  movel([0.339541, -0.797675, -2.797193, -1.117521, 1.570796, 1.910338],accel_mss,speed_ms,0,blend_radius_m)
  movel([0.338270, -0.798291, -2.797090, -1.117008, 1.570796, 1.909067],accel_mss,speed_ms,0,blend_radius_m)
  movel([0.337067, -0.798451, -2.797063, -1.116875, 1.570796, 1.907863],accel_mss,speed_ms,0,blend_radius_m)
  movel([0.336030, -0.798308, -2.797087, -1.116993, 1.570796, 1.906826],accel_mss,speed_ms,0,blend_radius_m)
  movel([0.330509, -0.796529, -2.797384, -1.118476, 1.570796, 1.901306],accel_mss,speed_ms,0,blend_radius_m)
  movel([0.325271, -0.794328, -2.797750, -1.120311, 1.570796, 1.896067],accel_mss,speed_ms,0,blend_radius_m)
  movel([0.320318, -0.791707, -2.798181, -1.122501, 1.570796, 1.891115],accel_mss,speed_ms,0,blend_radius_m)
  movel([0.315671, -0.788660, -2.798679, -1.125051, 1.570796, 1.886468],accel_mss,speed_ms,0,blend_radius_m)
  movel([0.314088, -0.787352, -2.798891, -1.126146, 1.570796, 1.884885],accel_mss,speed_ms,0,blend_radius_m)
  movel([0.312919, -0.785569, -2.799178, -1.127642, 1.570796, 1.883716],accel_mss,speed_ms,0,blend_radius_m)
  movel([0.312565, -0.784172, -2.799403, -1.128814, 1.570796, 1.883362],accel_mss,speed_ms,0,blend_radius_m)
  movel([0.312427, -0.782583, -2.799657, -1.130150, 1.570796, 1.883224],accel_mss,speed_ms,0,blend_radius_m)
  movel([0.312533, -0.779070, -2.800213, -1.133105, 1.570796, 1.883329],accel_mss,speed_ms,0,blend_radius_m)
  movel([0.314201, -0.765515, -2.802305, -1.144570, 1.570796, 1.884998],accel_mss,speed_ms,0,blend_radius_m)
  movel([0.314322, -0.761910, -2.802846, -1.147634, 1.570796, 1.885118],accel_mss,speed_ms,0,blend_radius_m)
  movel([0.313995, -0.758978, -2.803281, -1.150130, 1.570796, 1.884791],accel_mss,speed_ms,0,blend_radius_m)
  movel([0.313608, -0.757890, -2.803441, -1.151058, 1.570796, 1.884404],accel_mss,speed_ms,0,blend_radius_m)
  movel([0.313044, -0.757111, -2.803556, -1.151722, 1.570796, 1.883841],accel_mss,speed_ms,0,blend_radius_m)
  movel([0.312284, -0.756701, -2.803616, -1.152072, 1.570796, 1.883080],accel_mss,speed_ms,0,blend_radius_m)
  movel([0.311307, -0.756696, -2.803617, -1.152076, 1.570796, 1.882104],accel_mss,speed_ms,0,blend_radius_m)
  movel([0.309324, -0.757338, -2.803522, -1.151529, 1.570796, 1.880120],accel_mss,speed_ms,0,blend_radius_m)
  movel([0.308425, -0.757514, -2.803496, -1.151378, 1.570796, 1.879221],accel_mss,speed_ms,0,blend_radius_m)
  movel([0.307786, -0.757283, -2.803531, -1.151575, 1.570796, 1.878582],accel_mss,speed_ms,0,blend_radius_m)
  movel([0.307584, -0.756087, -2.803706, -1.152596, 1.570796, 1.878380],accel_mss,speed_ms,0,blend_radius_m)
  movel([0.307977, -0.754391, -2.803953, -1.154044, 1.570796, 1.878773],accel_mss,speed_ms,0,blend_radius_m)
  movel([0.309463, -0.748829, -2.804756, -1.158804, 1.570796, 1.880260],accel_mss,speed_ms,0,blend_radius_m)
  movel([0.310630, -0.743455, -2.805517, -1.163417, 1.570796, 1.881426],accel_mss,speed_ms,0,blend_radius_m)
  movel([0.312165, -0.733164, -2.806936, -1.172289, 1.570796, 1.882961],accel_mss,speed_ms,0,blend_radius_m)
  movel([0.312944, -0.723256, -2.808256, -1.180876, 1.570796, 1.883740],accel_mss,speed_ms,0,blend_radius_m)
  movel([0.313326, -0.713471, -2.809516, -1.189402, 1.570796, 1.884122],accel_mss,speed_ms,0,blend_radius_m)
  speed_ms = 0.005
  movel([0.313326, -0.706215, -2.802909, -1.203265, 1.570796, 1.884122],accel_mss,speed_ms,0,blend_radius_m)
  speed_ms = 0.040
  movel([0.305588, -0.724600, -2.800519, -1.187270, 1.570796, 1.876385],accel_mss,speed_ms,0,blend_radius_m)
  speed_ms = 0.005
  movel([0.305588, -0.732101, -2.807080, -1.173208, 1.570796, 1.876385],accel_mss,speed_ms,0,blend_radius_m)
  speed_ms = 0.025
  movel([0.301170, -0.744287, -2.805400, -1.162703, 1.570796, 1.871966],accel_mss,speed_ms,0,blend_radius_m)
  movel([0.298692, -0.750428, -2.804526, -1.157434, 1.570796, 1.869489],accel_mss,speed_ms,0,blend_radius_m)
  movel([0.296052, -0.756579, -2.803634, -1.152176, 1.570796, 1.866849],accel_mss,speed_ms,0,blend_radius_m)
  movel([0.293909, -0.755261, -2.803827, -1.153301, 1.570796, 1.864706],accel_mss,speed_ms,0,blend_radius_m)
  movel([0.293492, -0.755110, -2.803849, -1.153430, 1.570796, 1.864289],accel_mss,speed_ms,0,blend_radius_m)
  movel([0.292925, -0.755314, -2.803819, -1.153256, 1.570796, 1.863721],accel_mss,speed_ms,0,blend_radius_m)
  movel([0.292315, -0.755987, -2.803720, -1.152681, 1.570796, 1.863111],accel_mss,speed_ms,0,blend_radius_m)
  movel([0.291839, -0.756807, -2.803600, -1.151981, 1.570796, 1.862635],accel_mss,speed_ms,0,blend_radius_m)
  movel([0.288894, -0.761863, -2.802853, -1.147674, 1.570796, 1.859691],accel_mss,speed_ms,0,blend_radius_m)
  movel([0.285493, -0.766786, -2.802112, -1.143491, 1.570796, 1.856290],accel_mss,speed_ms,0,blend_radius_m)
  movel([0.284595, -0.767854, -2.801950, -1.142584, 1.570796, 1.855391],accel_mss,speed_ms,0,blend_radius_m)
  movel([0.283710, -0.768447, -2.801860, -1.142082, 1.570796, 1.854506],accel_mss,speed_ms,0,blend_radius_m)
  movel([0.283279, -0.768196, -2.801898, -1.142295, 1.570796, 1.854075],accel_mss,speed_ms,0,blend_radius_m)
  movel([0.283199, -0.767514, -2.802002, -1.142873, 1.570796, 1.853995],accel_mss,speed_ms,0,blend_radius_m)
  movel([0.283611, -0.762679, -2.802731, -1.146980, 1.570796, 1.854408],accel_mss,speed_ms,0,blend_radius_m)
  movel([0.284807, -0.757324, -2.803525, -1.151541, 1.570796, 1.855604],accel_mss,speed_ms,0,blend_radius_m)
  speed_ms = 0.005
  movel([0.284807, -0.749511, -2.797028, -1.165850, 1.570796, 1.855604],accel_mss,speed_ms,0,blend_radius_m)
  speed_ms = 0.040
  movel([0.290706, -0.756584, -2.795983, -1.159821, 1.570796, 1.861503],accel_mss,speed_ms,0,blend_radius_m)
  speed_ms = 0.005
  movel([0.290706, -0.764482, -2.802460, -1.145446, 1.570796, 1.861503],accel_mss,speed_ms,0,blend_radius_m)
  speed_ms = 0.025
  movel([0.289009, -0.772297, -2.801270, -1.138822, 1.570796, 1.859805],accel_mss,speed_ms,0,blend_radius_m)
  movel([0.287811, -0.776370, -2.800637, -1.135382, 1.570796, 1.858608],accel_mss,speed_ms,0,blend_radius_m)
  movel([0.284778, -0.784728, -2.799313, -1.128347, 1.570796, 1.855575],accel_mss,speed_ms,0,blend_radius_m)
  movel([0.282956, -0.788978, -2.798627, -1.124784, 1.570796, 1.853753],accel_mss,speed_ms,0,blend_radius_m)
  movel([0.278747, -0.797523, -2.797219, -1.117648, 1.570796, 1.849544],accel_mss,speed_ms,0,blend_radius_m)
  movel([0.279478, -0.794879, -2.797658, -1.119852, 1.570796, 1.850275],accel_mss,speed_ms,0,blend_radius_m)
  movel([0.279565, -0.792616, -2.798032, -1.121741, 1.570796, 1.850361],accel_mss,speed_ms,0,blend_radius_m)
  movel([0.279016, -0.790889, -2.798315, -1.123185, 1.570796, 1.849813],accel_mss,speed_ms,0,blend_radius_m)
  movel([0.277841, -0.789851, -2.798485, -1.124053, 1.570796, 1.848637],accel_mss,speed_ms,0,blend_radius_m)
  speed_ms = 0.005
  movel([0.277841, -0.781667, -2.792079, -1.138643, 1.570796, 1.848637],accel_mss,speed_ms,0,blend_radius_m)
  speed_ms = 0.040
  movel([0.251919, -0.798788, -2.789231, -1.124370, 1.570796, 1.822716],accel_mss,speed_ms,0,blend_radius_m)
  speed_ms = 0.005
  movel([0.251919, -0.807155, -2.795586, -1.109648, 1.570796, 1.822716],accel_mss,speed_ms,0,blend_radius_m)
  speed_ms = 0.025
  movel([0.247378, -0.813004, -2.794571, -1.104814, 1.570796, 1.818174],accel_mss,speed_ms,0,blend_radius_m)
  movel([0.242549, -0.818489, -2.793603, -1.100297, 1.570796, 1.813345],accel_mss,speed_ms,0,blend_radius_m)
  movel([0.237519, -0.823531, -2.792698, -1.096159, 1.570796, 1.808315],accel_mss,speed_ms,0,blend_radius_m)
  movel([0.232368, -0.828046, -2.791877, -1.092466, 1.570796, 1.803164],accel_mss,speed_ms,0,blend_radius_m)
  movel([0.233688, -0.825444, -2.792352, -1.094593, 1.570796, 1.804484],accel_mss,speed_ms,0,blend_radius_m)
  movel([0.234683, -0.823023, -2.792790, -1.096576, 1.570796, 1.805479],accel_mss,speed_ms,0,blend_radius_m)
  movel([0.235280, -0.821000, -2.793154, -1.098235, 1.570796, 1.806076],accel_mss,speed_ms,0,blend_radius_m)
  movel([0.235407, -0.819588, -2.793407, -1.099394, 1.570796, 1.806203],accel_mss,speed_ms,0,blend_radius_m)
  movel([0.234984, -0.819018, -2.793509, -1.099863, 1.570796, 1.805780],accel_mss,speed_ms,0,blend_radius_m)
  movel([0.234547, -0.819112, -2.793492, -1.099785, 1.570796, 1.805344],accel_mss,speed_ms,0,blend_radius_m)
  movel([0.233940, -0.819499, -2.793423, -1.099468, 1.570796, 1.804736],accel_mss,speed_ms,0,blend_radius_m)
  movel([0.232209, -0.821250, -2.793109, -1.098030, 1.570796, 1.803005],accel_mss,speed_ms,0,blend_radius_m)
  movel([0.227802, -0.827037, -2.792062, -1.093291, 1.570796, 1.798598],accel_mss,speed_ms,0,blend_radius_m)
  movel([0.225752, -0.829544, -2.791602, -1.091243, 1.570796, 1.796549],accel_mss,speed_ms,0,blend_radius_m)
  movel([0.221376, -0.834255, -2.790729, -1.087405, 1.570796, 1.792172],accel_mss,speed_ms,0,blend_radius_m)
  movel([0.219102, -0.836398, -2.790328, -1.085663, 1.570796, 1.789898],accel_mss,speed_ms,0,blend_radius_m)
  movel([0.216804, -0.838351, -2.789960, -1.084077, 1.570796, 1.787600],accel_mss,speed_ms,0,blend_radius_m)
  movel([0.214506, -0.840095, -2.789630, -1.082663, 1.570796, 1.785302],accel_mss,speed_ms,0,blend_radius_m)
  movel([0.212240, -0.841584, -2.789347, -1.081458, 1.570796, 1.783037],accel_mss,speed_ms,0,blend_radius_m)
  movel([0.215104, -0.837462, -2.790128, -1.084799, 1.570796, 1.785901],accel_mss,speed_ms,0,blend_radius_m)
  movel([0.217906, -0.833284, -2.790910, -1.088195, 1.570796, 1.788702],accel_mss,speed_ms,0,blend_radius_m)
  movel([0.219209, -0.830564, -2.791414, -1.090411, 1.570796, 1.790005],accel_mss,speed_ms,0,blend_radius_m)
  movel([0.219966, -0.827999, -2.791886, -1.092505, 1.570796, 1.790763],accel_mss,speed_ms,0,blend_radius_m)
  movel([0.219920, -0.827191, -2.792033, -1.093165, 1.570796, 1.790716],accel_mss,speed_ms,0,blend_radius_m)
  movel([0.219466, -0.826927, -2.792082, -1.093380, 1.570796, 1.790262],accel_mss,speed_ms,0,blend_radius_m)
  movel([0.218525, -0.827372, -2.792000, -1.093017, 1.570796, 1.789321],accel_mss,speed_ms,0,blend_radius_m)
  movel([0.217006, -0.828695, -2.791758, -1.091936, 1.570796, 1.787803],accel_mss,speed_ms,0,blend_radius_m)
  movel([0.209003, -0.836814, -2.790250, -1.085325, 1.570796, 1.779799],accel_mss,speed_ms,0,blend_radius_m)
  movel([0.205006, -0.840380, -2.789576, -1.082433, 1.570796, 1.775803],accel_mss,speed_ms,0,blend_radius_m)
  movel([0.203015, -0.841850, -2.789296, -1.081243, 1.570796, 1.773811],accel_mss,speed_ms,0,blend_radius_m)
  movel([0.201023, -0.843044, -2.789068, -1.080276, 1.570796, 1.771819],accel_mss,speed_ms,0,blend_radius_m)
  speed_ms = 0.005
  movel([0.201023, -0.834334, -2.782823, -1.095231, 1.570796, 1.771819],accel_mss,speed_ms,0,blend_radius_m)
  speed_ms = 0.040
  movel([0.238662, -0.779480, -2.792432, -1.140477, 1.570796, 1.809458],accel_mss,speed_ms,0,blend_radius_m)
  speed_ms = 0.005
  movel([0.238662, -0.787640, -2.798844, -1.125905, 1.570796, 1.809458],accel_mss,speed_ms,0,blend_radius_m)
  speed_ms = 0.025
  movel([0.238890, -0.784551, -2.799342, -1.128496, 1.570796, 1.809686],accel_mss,speed_ms,0,blend_radius_m)
  movel([0.239732, -0.781111, -2.799891, -1.131387, 1.570796, 1.810528],accel_mss,speed_ms,0,blend_radius_m)
  movel([0.241121, -0.777396, -2.800477, -1.134517, 1.570796, 1.811917],accel_mss,speed_ms,0,blend_radius_m)
  movel([0.242984, -0.773502, -2.801083, -1.137804, 1.570796, 1.813781],accel_mss,speed_ms,0,blend_radius_m)
  movel([0.245268, -0.769501, -2.801699, -1.141189, 1.570796, 1.816064],accel_mss,speed_ms,0,blend_radius_m)
  movel([0.247890, -0.765497, -2.802307, -1.144584, 1.570796, 1.818687],accel_mss,speed_ms,0,blend_radius_m)
  movel([0.250794, -0.761568, -2.802896, -1.147924, 1.570796, 1.821590],accel_mss,speed_ms,0,blend_radius_m)
  movel([0.253896, -0.757818, -2.803452, -1.151119, 1.570796, 1.824692],accel_mss,speed_ms,0,blend_radius_m)
  movel([0.257898, -0.753459, -2.804089, -1.154841, 1.570796, 1.828695],accel_mss,speed_ms,0,blend_radius_m)
  movel([0.266086, -0.744895, -2.805314, -1.162180, 1.570796, 1.836882],accel_mss,speed_ms,0,blend_radius_m)
  movel([0.270058, -0.740350, -2.805950, -1.166089, 1.570796, 1.840855],accel_mss,speed_ms,0,blend_radius_m)
  movel([0.273771, -0.735350, -2.806639, -1.170400, 1.570796, 1.844568],accel_mss,speed_ms,0,blend_radius_m)
  movel([0.275420, -0.732740, -2.806993, -1.172655, 1.570796, 1.846216],accel_mss,speed_ms,0,blend_radius_m)
  movel([0.276854, -0.730144, -2.807343, -1.174902, 1.570796, 1.847650],accel_mss,speed_ms,0,blend_radius_m)
  movel([0.278016, -0.727626, -2.807680, -1.177084, 1.570796, 1.848812],accel_mss,speed_ms,0,blend_radius_m)
  movel([0.278854, -0.725248, -2.807995, -1.179146, 1.570796, 1.849650],accel_mss,speed_ms,0,blend_radius_m)
  movel([0.279296, -0.723094, -2.808277, -1.181017, 1.570796, 1.850092],accel_mss,speed_ms,0,blend_radius_m)
  movel([0.279283, -0.721232, -2.808520, -1.182636, 1.570796, 1.850080],accel_mss,speed_ms,0,blend_radius_m)
  speed_ms = 0.005
  movel([0.279283, -0.713873, -2.801932, -1.196584, 1.570796, 1.850080],accel_mss,speed_ms,0,blend_radius_m)
  speed_ms = 0.040
  movel([0.278218, -0.699673, -2.803723, -1.208993, 1.570796, 1.849015],accel_mss,speed_ms,0,blend_radius_m)
  speed_ms = 0.005
  movel([0.278218, -0.706840, -2.810345, -1.195204, 1.570796, 1.849015],accel_mss,speed_ms,0,blend_radius_m)
  speed_ms = 0.025
  movel([0.274128, -0.720252, -2.808648, -1.183489, 1.570796, 1.844925],accel_mss,speed_ms,0,blend_radius_m)
  movel([0.272708, -0.723399, -2.808238, -1.180753, 1.570796, 1.843504],accel_mss,speed_ms,0,blend_radius_m)
  movel([0.270637, -0.726538, -2.807824, -1.178027, 1.570796, 1.841433],accel_mss,speed_ms,0,blend_radius_m)
  movel([0.268156, -0.729467, -2.807434, -1.175488, 1.570796, 1.838952],accel_mss,speed_ms,0,blend_radius_m)
  movel([0.259858, -0.738116, -2.806259, -1.168014, 1.570796, 1.830654],accel_mss,speed_ms,0,blend_radius_m)
  movel([0.257055, -0.741410, -2.805803, -1.165176, 1.570796, 1.827852],accel_mss,speed_ms,0,blend_radius_m)
  movel([0.254399, -0.744824, -2.805324, -1.162241, 1.570796, 1.825196],accel_mss,speed_ms,0,blend_radius_m)
  movel([0.251913, -0.748315, -2.804829, -1.159245, 1.570796, 1.822709],accel_mss,speed_ms,0,blend_radius_m)
  movel([0.249806, -0.751776, -2.804332, -1.156281, 1.570796, 1.820602],accel_mss,speed_ms,0,blend_radius_m)
  movel([0.248006, -0.755228, -2.803831, -1.153329, 1.570796, 1.818802],accel_mss,speed_ms,0,blend_radius_m)
  movel([0.246241, -0.758651, -2.803329, -1.150409, 1.570796, 1.817038],accel_mss,speed_ms,0,blend_radius_m)
  movel([0.244246, -0.762033, -2.802827, -1.147529, 1.570796, 1.815042],accel_mss,speed_ms,0,blend_radius_m)
  movel([0.242758, -0.756334, -2.803670, -1.152385, 1.570796, 1.813555],accel_mss,speed_ms,0,blend_radius_m)
  movel([0.243050, -0.754319, -2.803964, -1.154106, 1.570796, 1.813846],accel_mss,speed_ms,0,blend_radius_m)
  movel([0.243651, -0.752175, -2.804275, -1.155940, 1.570796, 1.814448],accel_mss,speed_ms,0,blend_radius_m)
  movel([0.244562, -0.749898, -2.804603, -1.157888, 1.570796, 1.815359],accel_mss,speed_ms,0,blend_radius_m)
  movel([0.245801, -0.747468, -2.804950, -1.159971, 1.570796, 1.816598],accel_mss,speed_ms,0,blend_radius_m)
  movel([0.248098, -0.744058, -2.805432, -1.162899, 1.570796, 1.818894],accel_mss,speed_ms,0,blend_radius_m)
  movel([0.251441, -0.739885, -2.806015, -1.166489, 1.570796, 1.822238],accel_mss,speed_ms,0,blend_radius_m)
  movel([0.259675, -0.730420, -2.807306, -1.174663, 1.570796, 1.830471],accel_mss,speed_ms,0,blend_radius_m)
  movel([0.263755, -0.725728, -2.807931, -1.178730, 1.570796, 1.834551],accel_mss,speed_ms,0,blend_radius_m)
  movel([0.267253, -0.721467, -2.808490, -1.182432, 1.570796, 1.838049],accel_mss,speed_ms,0,blend_radius_m)
  movel([0.269743, -0.717961, -2.808943, -1.185485, 1.570796, 1.840539],accel_mss,speed_ms,0,blend_radius_m)
  movel([0.270479, -0.716582, -2.809120, -1.186687, 1.570796, 1.841275],accel_mss,speed_ms,0,blend_radius_m)
  movel([0.270799, -0.715510, -2.809257, -1.187622, 1.570796, 1.841595],accel_mss,speed_ms,0,blend_radius_m)
  speed_ms = 0.005
  movel([0.270799, -0.708226, -2.802655, -1.201508, 1.570796, 1.841595],accel_mss,speed_ms,0,blend_radius_m)
  speed_ms = 0.040
  movel([0.256086, -0.711101, -2.802289, -1.198999, 1.570796, 1.826882],accel_mss,speed_ms,0,blend_radius_m)
  speed_ms = 0.005
  movel([0.256086, -0.718423, -2.808884, -1.185082, 1.570796, 1.826882],accel_mss,speed_ms,0,blend_radius_m)
  speed_ms = 0.025
  movel([0.254666, -0.718676, -2.808851, -1.184862, 1.570796, 1.825462],accel_mss,speed_ms,0,blend_radius_m)
  movel([0.253508, -0.718501, -2.808874, -1.185014, 1.570796, 1.824304],accel_mss,speed_ms,0,blend_radius_m)
  movel([0.251855, -0.717143, -2.809048, -1.186198, 1.570796, 1.822651],accel_mss,speed_ms,0,blend_radius_m)
  movel([0.250882, -0.714842, -2.809342, -1.188205, 1.570796, 1.821679],accel_mss,speed_ms,0,blend_radius_m)
  movel([0.250362, -0.712082, -2.809691, -1.190616, 1.570796, 1.821158],accel_mss,speed_ms,0,blend_radius_m)
  movel([0.250376, -0.710916, -2.809838, -1.191635, 1.570796, 1.821172],accel_mss,speed_ms,0,blend_radius_m)
  movel([0.251431, -0.708572, -2.810131, -1.193686, 1.570796, 1.822227],accel_mss,speed_ms,0,blend_radius_m)
  movel([0.255097, -0.701778, -2.810965, -1.199646, 1.570796, 1.825893],accel_mss,speed_ms,0,blend_radius_m)
  movel([0.261993, -0.688097, -2.812584, -1.211708, 1.570796, 1.832789],accel_mss,speed_ms,0,blend_radius_m)
  movel([0.265206, -0.681243, -2.813364, -1.217782, 1.570796, 1.836002],accel_mss,speed_ms,0,blend_radius_m)
  speed_ms = 0.005
  movel([0.265206, -0.674435, -2.806684, -1.231270, 1.570796, 1.836002],accel_mss,speed_ms,0,blend_radius_m)
  speed_ms = 0.040
  movel([0.255172, -0.681907, -2.805837, -1.224645, 1.570796, 1.825968],accel_mss,speed_ms,0,blend_radius_m)
  speed_ms = 0.005
  movel([0.255172, -0.688824, -2.812500, -1.211066, 1.570796, 1.825968],accel_mss,speed_ms,0,blend_radius_m)
  speed_ms = 0.025
  movel([0.253576, -0.692842, -2.812032, -1.207515, 1.570796, 1.824373],accel_mss,speed_ms,0,blend_radius_m)
  movel([0.251612, -0.696958, -2.811545, -1.203886, 1.570796, 1.822409],accel_mss,speed_ms,0,blend_radius_m)
  movel([0.249200, -0.700991, -2.811060, -1.200338, 1.570796, 1.819996],accel_mss,speed_ms,0,blend_radius_m)
  movel([0.247798, -0.702929, -2.810825, -1.198635, 1.570796, 1.818594],accel_mss,speed_ms,0,blend_radius_m)
  movel([0.244762, -0.706607, -2.810374, -1.195408, 1.570796, 1.815558],accel_mss,speed_ms,0,blend_radius_m)
  movel([0.243999, -0.708241, -2.810172, -1.193976, 1.570796, 1.814795],accel_mss,speed_ms,0,blend_radius_m)
  movel([0.239388, -0.720425, -2.808625, -1.183339, 1.570796, 1.810184],accel_mss,speed_ms,0,blend_radius_m)
  movel([0.238976, -0.721588, -2.808474, -1.182327, 1.570796, 1.809772],accel_mss,speed_ms,0,blend_radius_m)
  movel([0.238840, -0.722571, -2.808346, -1.181472, 1.570796, 1.809637],accel_mss,speed_ms,0,blend_radius_m)
  movel([0.239436, -0.723273, -2.808254, -1.180862, 1.570796, 1.810232],accel_mss,speed_ms,0,blend_radius_m)
  movel([0.240542, -0.723333, -2.808246, -1.180810, 1.570796, 1.811338],accel_mss,speed_ms,0,blend_radius_m)
  movel([0.243805, -0.723330, -2.808247, -1.180812, 1.570796, 1.814601],accel_mss,speed_ms,0,blend_radius_m)
  movel([0.246751, -0.723842, -2.808179, -1.180368, 1.570796, 1.817547],accel_mss,speed_ms,0,blend_radius_m)
  movel([0.249147, -0.725096, -2.808014, -1.179278, 1.570796, 1.819943],accel_mss,speed_ms,0,blend_radius_m)
  movel([0.250740, -0.727339, -2.807718, -1.177332, 1.570796, 1.821537],accel_mss,speed_ms,0,blend_radius_m)
  speed_ms = 0.005
  movel([0.250740, -0.719899, -2.801145, -1.191345, 1.570796, 1.821537],accel_mss,speed_ms,0,blend_radius_m)
  speed_ms = 0.040
  movel([0.239180, -0.750332, -2.796908, -1.165149, 1.570796, 1.809976],accel_mss,speed_ms,0,blend_radius_m)
  speed_ms = 0.005
  movel([0.239180, -0.758155, -2.803402, -1.150831, 1.570796, 1.809976],accel_mss,speed_ms,0,blend_radius_m)
  speed_ms = 0.025
  movel([0.238467, -0.758887, -2.803294, -1.150207, 1.570796, 1.809264],accel_mss,speed_ms,0,blend_radius_m)
  movel([0.237810, -0.759796, -2.803160, -1.149434, 1.570796, 1.808607],accel_mss,speed_ms,0,blend_radius_m)
  movel([0.235162, -0.764438, -2.802467, -1.145484, 1.570796, 1.805958],accel_mss,speed_ms,0,blend_radius_m)
  movel([0.234732, -0.764883, -2.802400, -1.145106, 1.570796, 1.805529],accel_mss,speed_ms,0,blend_radius_m)
  movel([0.234120, -0.765111, -2.802365, -1.144913, 1.570796, 1.804916],accel_mss,speed_ms,0,blend_radius_m)
  movel([0.233671, -0.764874, -2.802401, -1.145114, 1.570796, 1.804467],accel_mss,speed_ms,0,blend_radius_m)
  movel([0.233188, -0.763476, -2.802611, -1.146302, 1.570796, 1.803984],accel_mss,speed_ms,0,blend_radius_m)
  movel([0.233194, -0.760208, -2.803099, -1.149082, 1.570796, 1.803991],accel_mss,speed_ms,0,blend_radius_m)
  movel([0.234136, -0.756594, -2.803632, -1.152163, 1.570796, 1.804933],accel_mss,speed_ms,0,blend_radius_m)
  movel([0.235569, -0.752720, -2.804196, -1.155473, 1.570796, 1.806365],accel_mss,speed_ms,0,blend_radius_m)
  movel([0.237248, -0.748804, -2.804759, -1.158826, 1.570796, 1.808045],accel_mss,speed_ms,0,blend_radius_m)
  movel([0.239202, -0.744941, -2.805308, -1.162141, 1.570796, 1.809999],accel_mss,speed_ms,0,blend_radius_m)
  movel([0.241419, -0.741136, -2.805841, -1.165412, 1.570796, 1.812215],accel_mss,speed_ms,0,blend_radius_m)
  movel([0.243887, -0.737388, -2.806360, -1.168642, 1.570796, 1.814683],accel_mss,speed_ms,0,blend_radius_m)
  movel([0.246599, -0.733692, -2.806864, -1.171832, 1.570796, 1.817396],accel_mss,speed_ms,0,blend_radius_m)
  movel([0.249538, -0.730058, -2.807355, -1.174976, 1.570796, 1.820334],accel_mss,speed_ms,0,blend_radius_m)
  movel([0.252702, -0.726473, -2.807833, -1.178083, 1.570796, 1.823499],accel_mss,speed_ms,0,blend_radius_m)
  movel([0.256073, -0.722947, -2.808297, -1.181146, 1.570796, 1.826870],accel_mss,speed_ms,0,blend_radius_m)
  movel([0.260755, -0.717676, -2.808980, -1.185733, 1.570796, 1.831551],accel_mss,speed_ms,0,blend_radius_m)
  movel([0.265685, -0.711492, -2.809766, -1.191132, 1.570796, 1.836482],accel_mss,speed_ms,0,blend_radius_m)
  movel([0.271037, -0.704320, -2.810655, -1.197413, 1.570796, 1.841833],accel_mss,speed_ms,0,blend_radius_m)
  speed_ms = 0.005
  movel([0.271037, -0.697188, -2.804027, -1.211174, 1.570796, 1.841833],accel_mss,speed_ms,0,blend_radius_m)
  speed_ms = 0.040
  movel([0.266633, -0.698799, -2.803830, -1.209760, 1.570796, 1.837429],accel_mss,speed_ms,0,blend_radius_m)
  speed_ms = 0.005
  movel([0.266633, -0.705953, -2.810455, -1.195981, 1.570796, 1.837429],accel_mss,speed_ms,0,blend_radius_m)
  speed_ms = 0.025
  movel([0.271058, -0.696231, -2.811631, -1.204527, 1.570796, 1.841854],accel_mss,speed_ms,0,blend_radius_m)
  movel([0.275991, -0.686298, -2.812790, -1.213301, 1.570796, 1.846787],accel_mss,speed_ms,0,blend_radius_m)
  movel([0.278750, -0.681294, -2.813358, -1.217737, 1.570796, 1.849546],accel_mss,speed_ms,0,blend_radius_m)
  movel([0.281743, -0.676290, -2.813915, -1.222183, 1.570796, 1.852540],accel_mss,speed_ms,0,blend_radius_m)
  movel([0.285025, -0.671298, -2.814460, -1.226631, 1.570796, 1.855822],accel_mss,speed_ms,0,blend_radius_m)
  movel([0.288616, -0.666352, -2.814990, -1.231047, 1.570796, 1.859412],accel_mss,speed_ms,0,blend_radius_m)
  movel([0.298570, -0.653944, -2.816274, -1.242171, 1.570796, 1.869366],accel_mss,speed_ms,0,blend_radius_m)
  movel([0.302903, -0.648242, -2.816842, -1.247305, 1.570796, 1.873699],accel_mss,speed_ms,0,blend_radius_m)
  movel([0.304959, -0.645315, -2.817129, -1.249945, 1.570796, 1.875755],accel_mss,speed_ms,0,blend_radius_m)
  movel([0.306841, -0.642327, -2.817418, -1.252645, 1.570796, 1.877638],accel_mss,speed_ms,0,blend_radius_m)
  movel([0.311183, -0.633365, -2.818263, -1.260761, 1.570796, 1.881979],accel_mss,speed_ms,0,blend_radius_m)
  speed_ms = 0.005
  movel([0.311183, -0.627283, -2.811487, -1.273619, 1.570796, 1.881979],accel_mss,speed_ms,0,blend_radius_m)
  speed_ms = 0.040
  movel([0.321759, -0.606621, -2.813304, -1.292463, 1.570796, 1.892555],accel_mss,speed_ms,0,blend_radius_m)
  speed_ms = 0.005
  movel([0.321759, -0.612365, -2.820117, -1.279907, 1.570796, 1.892555],accel_mss,speed_ms,0,blend_radius_m)
  speed_ms = 0.025
  movel([0.325188, -0.604942, -2.820730, -1.286716, 1.570796, 1.895984],accel_mss,speed_ms,0,blend_radius_m)
  movel([0.327388, -0.601192, -2.821032, -1.290165, 1.570796, 1.898185],accel_mss,speed_ms,0,blend_radius_m)
  movel([0.330084, -0.597532, -2.821322, -1.293535, 1.570796, 1.900880],accel_mss,speed_ms,0,blend_radius_m)
  movel([0.332238, -0.595164, -2.821506, -1.295719, 1.570796, 1.903034],accel_mss,speed_ms,0,blend_radius_m)
  movel([0.334479, -0.593024, -2.821671, -1.297694, 1.570796, 1.905275],accel_mss,speed_ms,0,blend_radius_m)
  movel([0.339064, -0.589097, -2.821969, -1.301323, 1.570796, 1.909861],accel_mss,speed_ms,0,blend_radius_m)
  movel([0.343198, -0.585241, -2.822256, -1.304892, 1.570796, 1.913994],accel_mss,speed_ms,0,blend_radius_m)
  movel([0.346574, -0.581375, -2.822538, -1.308476, 1.570796, 1.917370],accel_mss,speed_ms,0,blend_radius_m)
  movel([0.353165, -0.572343, -2.823174, -1.316871, 1.570796, 1.923961],accel_mss,speed_ms,0,blend_radius_m)
  movel([0.354587, -0.570547, -2.823297, -1.318544, 1.570796, 1.925383],accel_mss,speed_ms,0,blend_radius_m)
  movel([0.356113, -0.568928, -2.823407, -1.320054, 1.570796, 1.926909],accel_mss,speed_ms,0,blend_radius_m)
  movel([0.359378, -0.566081, -2.823598, -1.322710, 1.570796, 1.930174],accel_mss,speed_ms,0,blend_radius_m)
  movel([0.365995, -0.560955, -2.823934, -1.327500, 1.570796, 1.936792],accel_mss,speed_ms,0,blend_radius_m)
  movel([0.373073, -0.554833, -2.824322, -1.333234, 1.570796, 1.943869],accel_mss,speed_ms,0,blend_radius_m)
  movel([0.376615, -0.551458, -2.824530, -1.336401, 1.570796, 1.947411],accel_mss,speed_ms,0,blend_radius_m)
  movel([0.380090, -0.547720, -2.824756, -1.339913, 1.570796, 1.950886],accel_mss,speed_ms,0,blend_radius_m)
  movel([0.382697, -0.544354, -2.824954, -1.343081, 1.570796, 1.953493],accel_mss,speed_ms,0,blend_radius_m)
  movel([0.384821, -0.540887, -2.825155, -1.346348, 1.570796, 1.955617],accel_mss,speed_ms,0,blend_radius_m)
  movel([0.385968, -0.537961, -2.825321, -1.349107, 1.570796, 1.956764],accel_mss,speed_ms,0,blend_radius_m)
  movel([0.386018, -0.536910, -2.825379, -1.350100, 1.570796, 1.956814],accel_mss,speed_ms,0,blend_radius_m)
  movel([0.385633, -0.536242, -2.825417, -1.350731, 1.570796, 1.956430],accel_mss,speed_ms,0,blend_radius_m)
  movel([0.384024, -0.535820, -2.825440, -1.351129, 1.570796, 1.954820],accel_mss,speed_ms,0,blend_radius_m)
  movel([0.381703, -0.536196, -2.825419, -1.350773, 1.570796, 1.952500],accel_mss,speed_ms,0,blend_radius_m)
  movel([0.378837, -0.537272, -2.825359, -1.349758, 1.570796, 1.949633],accel_mss,speed_ms,0,blend_radius_m)
  movel([0.375629, -0.538907, -2.825267, -1.348215, 1.570796, 1.946425],accel_mss,speed_ms,0,blend_radius_m)
  movel([0.372254, -0.541002, -2.825148, -1.346239, 1.570796, 1.943051],accel_mss,speed_ms,0,blend_radius_m)
  movel([0.368906, -0.543422, -2.825009, -1.343959, 1.570796, 1.939702],accel_mss,speed_ms,0,blend_radius_m)
  movel([0.365765, -0.546056, -2.824854, -1.341478, 1.570796, 1.936562],accel_mss,speed_ms,0,blend_radius_m)
  movel([0.363011, -0.548786, -2.824692, -1.338911, 1.570796, 1.933807],accel_mss,speed_ms,0,blend_radius_m)
  movel([0.359228, -0.553381, -2.824412, -1.334596, 1.570796, 1.930024],accel_mss,speed_ms,0,blend_radius_m)
  movel([0.348676, -0.567496, -2.823503, -1.321389, 1.570796, 1.919472],accel_mss,speed_ms,0,blend_radius_m)
  movel([0.341420, -0.576528, -2.822883, -1.312977, 1.570796, 1.912216],accel_mss,speed_ms,0,blend_radius_m)
  movel([0.334837, -0.583796, -2.822362, -1.306231, 1.570796, 1.905633],accel_mss,speed_ms,0,blend_radius_m)
  movel([0.331585, -0.587318, -2.822102, -1.302969, 1.570796, 1.902381],accel_mss,speed_ms,0,blend_radius_m)
  movel([0.328499, -0.590976, -2.821827, -1.299586, 1.570796, 1.899296],accel_mss,speed_ms,0,blend_radius_m)
  movel([0.325566, -0.594946, -2.821523, -1.295920, 1.570796, 1.896362],accel_mss,speed_ms,0,blend_radius_m)
  movel([0.322921, -0.598937, -2.821211, -1.292241, 1.570796, 1.893717],accel_mss,speed_ms,0,blend_radius_m)
  movel([0.320533, -0.602936, -2.820893, -1.288561, 1.570796, 1.891330],accel_mss,speed_ms,0,blend_radius_m)
  movel([0.318373, -0.606911, -2.820570, -1.284908, 1.570796, 1.889170],accel_mss,speed_ms,0,blend_radius_m)
  movel([0.314600, -0.614729, -2.819917, -1.277743, 1.570796, 1.885397],accel_mss,speed_ms,0,blend_radius_m)
  movel([0.311326, -0.622247, -2.819266, -1.270876, 1.570796, 1.882122],accel_mss,speed_ms,0,blend_radius_m)
  speed_ms = 0.005
  movel([0.311326, -0.616343, -2.812471, -1.283575, 1.570796, 1.882122],accel_mss,speed_ms,0,blend_radius_m)
  speed_ms = 0.040
  movel([0.303174, -0.623517, -2.811831, -1.277041, 1.570796, 1.873970],accel_mss,speed_ms,0,blend_radius_m)
  speed_ms = 0.005
  movel([0.303174, -0.629538, -2.818614, -1.264237, 1.570796, 1.873970],accel_mss,speed_ms,0,blend_radius_m)
  speed_ms = 0.025
  movel([0.308567, -0.617650, -2.819667, -1.275073, 1.570796, 1.879363],accel_mss,speed_ms,0,blend_radius_m)
  movel([0.311017, -0.612601, -2.820097, -1.279692, 1.570796, 1.881813],accel_mss,speed_ms,0,blend_radius_m)
  movel([0.313262, -0.607608, -2.820512, -1.284269, 1.570796, 1.884058],accel_mss,speed_ms,0,blend_radius_m)
  movel([0.314771, -0.603470, -2.820849, -1.288069, 1.570796, 1.885567],accel_mss,speed_ms,0,blend_radius_m)
  movel([0.315798, -0.599597, -2.821159, -1.291633, 1.570796, 1.886594],accel_mss,speed_ms,0,blend_radius_m)
  movel([0.316319, -0.596066, -2.821436, -1.294887, 1.570796, 1.887116],accel_mss,speed_ms,0,blend_radius_m)
  movel([0.316316, -0.592963, -2.821676, -1.297751, 1.570796, 1.887112],accel_mss,speed_ms,0,blend_radius_m)
  movel([0.318007, -0.591634, -2.821777, -1.298978, 1.570796, 1.888803],accel_mss,speed_ms,0,blend_radius_m)
  movel([0.319623, -0.590705, -2.821848, -1.299836, 1.570796, 1.890419],accel_mss,speed_ms,0,blend_radius_m)
  movel([0.322733, -0.589352, -2.821950, -1.301087, 1.570796, 1.893529],accel_mss,speed_ms,0,blend_radius_m)
  movel([0.326035, -0.587632, -2.822079, -1.302678, 1.570796, 1.896831],accel_mss,speed_ms,0,blend_radius_m)
  movel([0.327738, -0.586341, -2.822175, -1.303874, 1.570796, 1.898535],accel_mss,speed_ms,0,blend_radius_m)
  movel([0.329386, -0.584617, -2.822302, -1.305470, 1.570796, 1.900182],accel_mss,speed_ms,0,blend_radius_m)
  movel([0.348272, -0.561777, -2.823880, -1.326732, 1.570796, 1.919069],accel_mss,speed_ms,0,blend_radius_m)
  movel([0.348583, -0.559341, -2.824037, -1.329011, 1.570796, 1.919380],accel_mss,speed_ms,0,blend_radius_m)
  movel([0.348124, -0.557514, -2.824154, -1.330722, 1.570796, 1.918921],accel_mss,speed_ms,0,blend_radius_m)
  movel([0.346919, -0.556394, -2.824224, -1.331771, 1.570796, 1.917716],accel_mss,speed_ms,0,blend_radius_m)
  movel([0.345019, -0.556063, -2.824245, -1.332082, 1.570796, 1.915815],accel_mss,speed_ms,0,blend_radius_m)
  movel([0.348929, -0.553661, -2.824395, -1.334333, 1.570796, 1.919726],accel_mss,speed_ms,0,blend_radius_m)
  movel([0.352511, -0.552083, -2.824492, -1.335815, 1.570796, 1.923308],accel_mss,speed_ms,0,blend_radius_m)
  movel([0.355579, -0.551396, -2.824534, -1.336459, 1.570796, 1.926375],accel_mss,speed_ms,0,blend_radius_m)
  movel([0.357960, -0.551659, -2.824518, -1.336213, 1.570796, 1.928756],accel_mss,speed_ms,0,blend_radius_m)
  speed_ms = 0.005
  movel([0.357960, -0.546959, -2.817616, -1.347814, 1.570796, 1.928756],accel_mss,speed_ms,0,blend_radius_m)
  speed_ms = 0.040
  movel([0.361776, -0.536348, -2.818242, -1.357799, 1.570796, 1.932572],accel_mss,speed_ms,0,blend_radius_m)
  speed_ms = 0.005
  movel([0.361776, -0.540853, -2.825157, -1.346379, 1.570796, 1.932572],accel_mss,speed_ms,0,blend_radius_m)
  speed_ms = 0.025
  movel([0.364576, -0.534803, -2.825496, -1.352090, 1.570796, 1.935373],accel_mss,speed_ms,0,blend_radius_m)
  movel([0.366892, -0.529158, -2.825801, -1.357431, 1.570796, 1.937688],accel_mss,speed_ms,0,blend_radius_m)
  movel([0.368755, -0.523873, -2.826075, -1.362440, 1.570796, 1.939551],accel_mss,speed_ms,0,blend_radius_m)
  movel([0.370195, -0.518907, -2.826324, -1.367157, 1.570796, 1.940991],accel_mss,speed_ms,0,blend_radius_m)
  movel([0.371243, -0.514211, -2.826552, -1.371626, 1.570796, 1.942039],accel_mss,speed_ms,0,blend_radius_m)
  movel([0.371933, -0.509733, -2.826762, -1.375895, 1.570796, 1.942730],accel_mss,speed_ms,0,blend_radius_m)
  movel([0.372379, -0.501239, -2.827140, -1.384011, 1.570796, 1.943176],accel_mss,speed_ms,0,blend_radius_m)
  movel([0.362866, -0.522100, -2.826165, -1.364123, 1.570796, 1.933663],accel_mss,speed_ms,0,blend_radius_m)
  movel([0.363724, -0.519887, -2.826276, -1.366226, 1.570796, 1.934521],accel_mss,speed_ms,0,blend_radius_m)
  movel([0.364223, -0.517895, -2.826374, -1.368119, 1.570796, 1.935019],accel_mss,speed_ms,0,blend_radius_m)
  movel([0.364264, -0.514545, -2.826536, -1.371308, 1.570796, 1.935060],accel_mss,speed_ms,0,blend_radius_m)
  movel([0.363219, -0.511984, -2.826657, -1.373748, 1.570796, 1.934016],accel_mss,speed_ms,0,blend_radius_m)
  movel([0.361350, -0.510136, -2.826743, -1.375510, 1.570796, 1.932147],accel_mss,speed_ms,0,blend_radius_m)
  movel([0.358908, -0.508913, -2.826799, -1.376677, 1.570796, 1.929705],accel_mss,speed_ms,0,blend_radius_m)
  movel([0.356160, -0.508231, -2.826830, -1.377328, 1.570796, 1.926956],accel_mss,speed_ms,0,blend_radius_m)
  movel([0.350805, -0.508112, -2.826836, -1.377441, 1.570796, 1.921601],accel_mss,speed_ms,0,blend_radius_m)
  movel([0.352322, -0.514121, -2.826556, -1.371712, 1.570796, 1.923118],accel_mss,speed_ms,0,blend_radius_m)
  movel([0.352350, -0.517881, -2.826375, -1.368133, 1.570796, 1.923146],accel_mss,speed_ms,0,blend_radius_m)
  movel([0.351411, -0.522134, -2.826164, -1.364091, 1.570796, 1.922207],accel_mss,speed_ms,0,blend_radius_m)
  movel([0.349024, -0.523001, -2.826120, -1.363268, 1.570796, 1.919820],accel_mss,speed_ms,0,blend_radius_m)
  movel([0.346872, -0.523344, -2.826102, -1.362943, 1.570796, 1.917668],accel_mss,speed_ms,0,blend_radius_m)
  movel([0.342914, -0.523164, -2.826111, -1.363113, 1.570796, 1.913711],accel_mss,speed_ms,0,blend_radius_m)
  movel([0.338862, -0.522980, -2.826121, -1.363288, 1.570796, 1.909658],accel_mss,speed_ms,0,blend_radius_m)
  movel([0.336592, -0.523316, -2.826104, -1.362969, 1.570796, 1.907388],accel_mss,speed_ms,0,blend_radius_m)
  movel([0.334061, -0.524153, -2.826061, -1.362175, 1.570796, 1.904857],accel_mss,speed_ms,0,blend_radius_m)
  movel([0.331141, -0.529683, -2.825773, -1.356933, 1.570796, 1.901938],accel_mss,speed_ms,0,blend_radius_m)
  movel([0.329142, -0.534804, -2.825496, -1.352089, 1.570796, 1.899939],accel_mss,speed_ms,0,blend_radius_m)
  movel([0.325579, -0.536459, -2.825404, -1.350525, 1.570796, 1.896375],accel_mss,speed_ms,0,blend_radius_m)
  movel([0.322366, -0.537405, -2.825352, -1.349632, 1.570796, 1.893163],accel_mss,speed_ms,0,blend_radius_m)
  movel([0.319565, -0.537623, -2.825339, -1.349426, 1.570796, 1.890361],accel_mss,speed_ms,0,blend_radius_m)
  movel([0.317254, -0.537105, -2.825368, -1.349915, 1.570796, 1.888051],accel_mss,speed_ms,0,blend_radius_m)
  movel([0.316801, -0.537707, -2.825335, -1.349347, 1.570796, 1.887598],accel_mss,speed_ms,0,blend_radius_m)
  movel([0.312948, -0.544623, -2.824939, -1.342827, 1.570796, 1.883744],accel_mss,speed_ms,0,blend_radius_m)
  movel([0.308518, -0.553115, -2.824428, -1.334846, 1.570796, 1.879314],accel_mss,speed_ms,0,blend_radius_m)
  movel([0.306832, -0.557047, -2.824183, -1.331159, 1.570796, 1.877628],accel_mss,speed_ms,0,blend_radius_m)
  movel([0.305575, -0.560550, -2.823960, -1.327880, 1.570796, 1.876371],accel_mss,speed_ms,0,blend_radius_m)
  movel([0.303731, -0.567410, -2.823509, -1.321469, 1.570796, 1.874527],accel_mss,speed_ms,0,blend_radius_m)
  movel([0.296179, -0.564041, -2.823733, -1.324615, 1.570796, 1.866975],accel_mss,speed_ms,0,blend_radius_m)
  movel([0.294293, -0.568200, -2.823456, -1.320733, 1.570796, 1.865090],accel_mss,speed_ms,0,blend_radius_m)
  movel([0.292708, -0.572248, -2.823181, -1.316960, 1.570796, 1.863505],accel_mss,speed_ms,0,blend_radius_m)
  movel([0.290333, -0.579974, -2.822639, -1.309776, 1.570796, 1.861129],accel_mss,speed_ms,0,blend_radius_m)
  movel([0.288921, -0.587059, -2.822121, -1.303209, 1.570796, 1.859717],accel_mss,speed_ms,0,blend_radius_m)
  movel([0.288123, -0.595291, -2.821496, -1.295602, 1.570796, 1.858919],accel_mss,speed_ms,0,blend_radius_m)
  movel([0.287779, -0.596392, -2.821411, -1.294586, 1.570796, 1.858575],accel_mss,speed_ms,0,blend_radius_m)
  movel([0.287159, -0.597593, -2.821317, -1.293479, 1.570796, 1.857956],accel_mss,speed_ms,0,blend_radius_m)
  movel([0.285929, -0.599182, -2.821192, -1.292015, 1.570796, 1.856725],accel_mss,speed_ms,0,blend_radius_m)
  movel([0.276804, -0.608154, -2.820467, -1.283767, 1.570796, 1.847600],accel_mss,speed_ms,0,blend_radius_m)
  movel([0.272177, -0.612109, -2.820138, -1.280142, 1.570796, 1.842973],accel_mss,speed_ms,0,blend_radius_m)
  movel([0.270488, -0.613179, -2.820048, -1.279162, 1.570796, 1.841284],accel_mss,speed_ms,0,blend_radius_m)
  movel([0.269521, -0.613284, -2.820039, -1.279066, 1.570796, 1.840317],accel_mss,speed_ms,0,blend_radius_m)
  movel([0.273197, -0.615557, -2.819846, -1.276986, 1.570796, 1.843994],accel_mss,speed_ms,0,blend_radius_m)
  movel([0.275377, -0.616224, -2.819789, -1.276376, 1.570796, 1.846174],accel_mss,speed_ms,0,blend_radius_m)
  movel([0.277763, -0.616583, -2.819758, -1.276048, 1.570796, 1.848560],accel_mss,speed_ms,0,blend_radius_m)
  movel([0.269994, -0.626706, -2.818869, -1.266813, 1.570796, 1.840790],accel_mss,speed_ms,0,blend_radius_m)
  movel([0.261856, -0.637824, -2.817846, -1.256719, 1.570796, 1.832652],accel_mss,speed_ms,0,blend_radius_m)
  movel([0.258032, -0.643424, -2.817312, -1.251653, 1.570796, 1.828829],accel_mss,speed_ms,0,blend_radius_m)
  movel([0.254566, -0.648872, -2.816780, -1.246737, 1.570796, 1.825362],accel_mss,speed_ms,0,blend_radius_m)
  movel([0.251604, -0.654050, -2.816263, -1.242076, 1.570796, 1.822400],accel_mss,speed_ms,0,blend_radius_m)
  movel([0.249284, -0.658827, -2.815776, -1.237786, 1.570796, 1.820080],accel_mss,speed_ms,0,blend_radius_m)
  movel([0.252859, -0.655063, -2.816161, -1.241166, 1.570796, 1.823656],accel_mss,speed_ms,0,blend_radius_m)
  movel([0.256515, -0.651592, -2.816510, -1.244287, 1.570796, 1.827311],accel_mss,speed_ms,0,blend_radius_m)
  movel([0.260205, -0.648492, -2.816817, -1.247080, 1.570796, 1.831001],accel_mss,speed_ms,0,blend_radius_m)
  movel([0.263905, -0.645825, -2.817079, -1.249485, 1.570796, 1.834702],accel_mss,speed_ms,0,blend_radius_m)
  movel([0.261399, -0.648855, -2.816782, -1.246752, 1.570796, 1.832196],accel_mss,speed_ms,0,blend_radius_m)
  movel([0.256818, -0.655143, -2.816152, -1.241093, 1.570796, 1.827614],accel_mss,speed_ms,0,blend_radius_m)
  movel([0.254774, -0.658350, -2.815825, -1.238214, 1.570796, 1.825570],accel_mss,speed_ms,0,blend_radius_m)
  movel([0.251273, -0.664712, -2.815163, -1.232514, 1.570796, 1.822070],accel_mss,speed_ms,0,blend_radius_m)
  movel([0.249845, -0.667818, -2.814834, -1.229737, 1.570796, 1.820641],accel_mss,speed_ms,0,blend_radius_m)
  movel([0.248659, -0.670828, -2.814511, -1.227049, 1.570796, 1.819455],accel_mss,speed_ms,0,blend_radius_m)
  speed_ms = 0.005
  movel([0.248659, -0.664173, -2.807809, -1.240407, 1.570796, 1.819455],accel_mss,speed_ms,0,blend_radius_m)
  speed_ms = 0.040
  movel([0.261096, -0.665372, -2.807680, -1.239337, 1.570796, 1.831893],accel_mss,speed_ms,0,blend_radius_m)
  speed_ms = 0.005
  movel([0.261096, -0.672045, -2.814379, -1.225964, 1.570796, 1.831893],accel_mss,speed_ms,0,blend_radius_m)
  speed_ms = 0.025
  movel([0.261978, -0.668266, -2.814786, -1.229337, 1.570796, 1.832775],accel_mss,speed_ms,0,blend_radius_m)
  movel([0.263180, -0.664263, -2.815211, -1.232915, 1.570796, 1.833976],accel_mss,speed_ms,0,blend_radius_m)
  movel([0.264694, -0.660073, -2.815648, -1.236669, 1.570796, 1.835491],accel_mss,speed_ms,0,blend_radius_m)
  movel([0.266514, -0.655739, -2.816092, -1.240558, 1.570796, 1.837310],accel_mss,speed_ms,0,blend_radius_m)
  movel([0.268640, -0.651292, -2.816540, -1.244558, 1.570796, 1.839436],accel_mss,speed_ms,0,blend_radius_m)
  movel([0.271058, -0.646774, -2.816986, -1.248629, 1.570796, 1.841854],accel_mss,speed_ms,0,blend_radius_m)
  movel([0.273763, -0.642220, -2.817428, -1.252741, 1.570796, 1.844560],accel_mss,speed_ms,0,blend_radius_m)
  movel([0.276750, -0.637674, -2.817860, -1.256854, 1.570796, 1.847547],accel_mss,speed_ms,0,blend_radius_m)
  movel([0.286612, -0.623519, -2.819154, -1.269716, 1.570796, 1.857408],accel_mss,speed_ms,0,blend_radius_m)
  movel([0.288661, -0.620204, -2.819445, -1.272740, 1.570796, 1.859457],accel_mss,speed_ms,0,blend_radius_m)
  movel([0.290516, -0.616811, -2.819739, -1.275839, 1.570796, 1.861312],accel_mss,speed_ms,0,blend_radius_m)
  movel([0.292163, -0.613266, -2.820041, -1.279082, 1.570796, 1.862959],accel_mss,speed_ms,0,blend_radius_m)
  movel([0.293595, -0.609474, -2.820358, -1.282557, 1.570796, 1.864391],accel_mss,speed_ms,0,blend_radius_m)
  movel([0.296721, -0.598988, -2.821207, -1.292194, 1.570796, 1.867517],accel_mss,speed_ms,0,blend_radius_m)
  movel([0.298529, -0.593618, -2.821625, -1.297145, 1.570796, 1.869326],accel_mss,speed_ms,0,blend_radius_m)
  movel([0.301036, -0.587913, -2.822058, -1.302419, 1.570796, 1.871832],accel_mss,speed_ms,0,blend_radius_m)
  movel([0.303004, -0.584308, -2.822324, -1.305756, 1.570796, 1.873800],accel_mss,speed_ms,0,blend_radius_m)
  movel([0.305252, -0.580681, -2.822588, -1.309120, 1.570796, 1.876048],accel_mss,speed_ms,0,blend_radius_m)
  movel([0.310421, -0.573414, -2.823101, -1.315875, 1.570796, 1.881218],accel_mss,speed_ms,0,blend_radius_m)
  movel([0.316191, -0.566190, -2.823591, -1.322608, 1.570796, 1.886988],accel_mss,speed_ms,0,blend_radius_m)
  movel([0.322221, -0.559091, -2.824053, -1.329245, 1.570796, 1.893018],accel_mss,speed_ms,0,blend_radius_m)
  movel([0.328174, -0.552308, -2.824478, -1.335603, 1.570796, 1.898970],accel_mss,speed_ms,0,blend_radius_m)
  movel([0.334338, -0.545808, -2.824869, -1.341712, 1.570796, 1.905134],accel_mss,speed_ms,0,blend_radius_m)
  movel([0.337426, -0.542873, -2.825040, -1.344475, 1.570796, 1.908222],accel_mss,speed_ms,0,blend_radius_m)
  movel([0.340487, -0.540248, -2.825191, -1.346950, 1.570796, 1.911284],accel_mss,speed_ms,0,blend_radius_m)
  movel([0.343472, -0.538035, -2.825316, -1.349037, 1.570796, 1.914269],accel_mss,speed_ms,0,blend_radius_m)
  movel([0.346372, -0.536298, -2.825413, -1.350677, 1.570796, 1.917168],accel_mss,speed_ms,0,blend_radius_m)
  speed_ms = 0.005
  movel([0.346372, -0.531876, -2.818493, -1.362019, 1.570796, 1.917168],accel_mss,speed_ms,0,blend_radius_m)
  speed_ms = 0.040
  movel([0.349211, -0.533375, -2.818410, -1.360604, 1.570796, 1.920007],accel_mss,speed_ms,0,blend_radius_m)
  speed_ms = 0.005
  movel([0.349211, -0.537825, -2.825328, -1.349236, 1.570796, 1.920007],accel_mss,speed_ms,0,blend_radius_m)
  speed_ms = 0.025
  movel([0.350136, -0.538161, -2.825309, -1.348919, 1.570796, 1.920932],accel_mss,speed_ms,0,blend_radius_m)
  movel([0.351314, -0.538938, -2.825266, -1.348186, 1.570796, 1.922110],accel_mss,speed_ms,0,blend_radius_m)
  movel([0.352745, -0.542119, -2.825084, -1.345185, 1.570796, 1.923541],accel_mss,speed_ms,0,blend_radius_m)
  movel([0.352995, -0.544206, -2.824963, -1.343220, 1.570796, 1.923791],accel_mss,speed_ms,0,blend_radius_m)
  movel([0.352756, -0.545471, -2.824889, -1.342029, 1.570796, 1.923552],accel_mss,speed_ms,0,blend_radius_m)
  movel([0.352424, -0.545878, -2.824865, -1.341646, 1.570796, 1.923220],accel_mss,speed_ms,0,blend_radius_m)
  movel([0.351896, -0.546033, -2.824856, -1.341500, 1.570796, 1.922692],accel_mss,speed_ms,0,blend_radius_m)
  movel([0.346949, -0.545728, -2.824874, -1.341787, 1.570796, 1.917745],accel_mss,speed_ms,0,blend_radius_m)
  movel([0.344047, -0.546273, -2.824842, -1.341274, 1.570796, 1.914843],accel_mss,speed_ms,0,blend_radius_m)
  movel([0.342393, -0.547000, -2.824798, -1.340591, 1.570796, 1.913189],accel_mss,speed_ms,0,blend_radius_m)
  movel([0.340568, -0.548120, -2.824732, -1.339537, 1.570796, 1.911364],accel_mss,speed_ms,0,blend_radius_m)
  movel([0.338416, -0.549848, -2.824628, -1.337913, 1.570796, 1.909212],accel_mss,speed_ms,0,blend_radius_m)
  movel([0.336248, -0.551866, -2.824505, -1.336018, 1.570796, 1.907045],accel_mss,speed_ms,0,blend_radius_m)
  movel([0.330981, -0.557235, -2.824171, -1.330983, 1.570796, 1.901778],accel_mss,speed_ms,0,blend_radius_m)
  movel([0.325797, -0.563012, -2.823800, -1.325577, 1.570796, 1.896593],accel_mss,speed_ms,0,blend_radius_m)
  movel([0.320854, -0.569013, -2.823401, -1.319974, 1.570796, 1.891650],accel_mss,speed_ms,0,blend_radius_m)
  movel([0.316321, -0.575033, -2.822988, -1.314368, 1.570796, 1.887118],accel_mss,speed_ms,0,blend_radius_m)
  movel([0.318210, -0.579379, -2.822681, -1.310328, 1.570796, 1.889007],accel_mss,speed_ms,0,blend_radius_m)
  movel([0.319268, -0.584570, -2.822305, -1.305514, 1.570796, 1.890065],accel_mss,speed_ms,0,blend_radius_m)
  movel([0.317463, -0.584332, -2.822323, -1.305734, 1.570796, 1.888260],accel_mss,speed_ms,0,blend_radius_m)
  movel([0.315279, -0.584721, -2.822294, -1.305374, 1.570796, 1.886076],accel_mss,speed_ms,0,blend_radius_m)
  movel([0.312783, -0.585732, -2.822220, -1.304437, 1.570796, 1.883579],accel_mss,speed_ms,0,blend_radius_m)
  movel([0.310067, -0.587325, -2.822101, -1.302962, 1.570796, 1.880864],accel_mss,speed_ms,0,blend_radius_m)
  movel([0.308732, -0.588520, -2.822012, -1.301857, 1.570796, 1.879528],accel_mss,speed_ms,0,blend_radius_m)
  movel([0.308074, -0.589870, -2.821911, -1.300608, 1.570796, 1.878870],accel_mss,speed_ms,0,blend_radius_m)
  movel([0.303568, -0.603434, -2.820852, -1.288103, 1.570796, 1.874364],accel_mss,speed_ms,0,blend_radius_m)
  movel([0.300842, -0.610507, -2.820272, -1.281610, 1.570796, 1.871639],accel_mss,speed_ms,0,blend_radius_m)
  movel([0.297673, -0.617839, -2.819650, -1.274900, 1.570796, 1.868470],accel_mss,speed_ms,0,blend_radius_m)
  movel([0.294091, -0.625251, -2.819000, -1.268138, 1.570796, 1.864887],accel_mss,speed_ms,0,blend_radius_m)
  movel([0.290108, -0.632581, -2.818335, -1.261473, 1.570796, 1.860904],accel_mss,speed_ms,0,blend_radius_m)
  movel([0.281824, -0.647250, -2.816940, -1.248199, 1.570796, 1.852621],accel_mss,speed_ms,0,blend_radius_m)
  movel([0.278355, -0.654316, -2.816236, -1.241837, 1.570796, 1.849151],accel_mss,speed_ms,0,blend_radius_m)
  movel([0.275692, -0.661168, -2.815534, -1.235687, 1.570796, 1.846488],accel_mss,speed_ms,0,blend_radius_m)
  speed_ms = 0.005
  movel([0.275692, -0.654656, -2.808812, -1.248921, 1.570796, 1.846488],accel_mss,speed_ms,0,blend_radius_m)
  speed_ms = 0.040
  movel([0.303078, -0.634872, -2.810777, -1.266740, 1.570796, 1.873874],accel_mss,speed_ms,0,blend_radius_m)
  speed_ms = 0.005
  movel([0.303078, -0.641076, -2.817538, -1.253775, 1.570796, 1.873874],accel_mss,speed_ms,0,blend_radius_m)
  speed_ms = 0.025
  movel([0.300877, -0.646685, -2.816995, -1.248709, 1.570796, 1.871673],accel_mss,speed_ms,0,blend_radius_m)
  movel([0.297944, -0.652518, -2.816417, -1.243454, 1.570796, 1.868740],accel_mss,speed_ms,0,blend_radius_m)
  movel([0.294388, -0.658376, -2.815823, -1.238191, 1.570796, 1.865184],accel_mss,speed_ms,0,blend_radius_m)
  movel([0.290325, -0.664072, -2.815231, -1.233086, 1.570796, 1.861122],accel_mss,speed_ms,0,blend_radius_m)
  speed_ms = 0.005
  movel([0.290325, -0.657517, -2.808515, -1.246357, 1.570796, 1.861122],accel_mss,speed_ms,0,blend_radius_m)
  speed_ms = 0.040
  movel([0.285559, -0.653551, -2.808926, -1.249911, 1.570796, 1.856356],accel_mss,speed_ms,0,blend_radius_m)
  speed_ms = 0.005
  movel([0.285559, -0.660046, -2.815650, -1.236692, 1.570796, 1.856356],accel_mss,speed_ms,0,blend_radius_m)
  speed_ms = 0.025
  movel([0.265122, -0.696171, -2.811638, -1.204580, 1.570796, 1.835919],accel_mss,speed_ms,0,blend_radius_m)
  movel([0.264110, -0.698390, -2.811374, -1.202626, 1.570796, 1.834906],accel_mss,speed_ms,0,blend_radius_m)
  movel([0.264152, -0.700398, -2.811132, -1.200859, 1.570796, 1.834948],accel_mss,speed_ms,0,blend_radius_m)
  movel([0.264198, -0.702992, -2.810817, -1.198580, 1.570796, 1.834995],accel_mss,speed_ms,0,blend_radius_m)
  movel([0.263580, -0.706069, -2.810440, -1.195880, 1.570796, 1.834376],accel_mss,speed_ms,0,blend_radius_m)
  speed_ms = 0.005
  movel([0.263580, -0.698913, -2.803816, -1.209660, 1.570796, 1.834376],accel_mss,speed_ms,0,blend_radius_m)
  speed_ms = 0.040
  movel([0.294514, -0.672200, -2.806933, -1.233256, 1.570796, 1.865311],accel_mss,speed_ms,0,blend_radius_m)
  speed_ms = 0.005
  movel([0.294514, -0.678975, -2.813618, -1.219796, 1.570796, 1.865311],accel_mss,speed_ms,0,blend_radius_m)
  speed_ms = 0.025
  movel([0.295315, -0.675586, -2.813993, -1.222810, 1.570796, 1.866111],accel_mss,speed_ms,0,blend_radius_m)
  movel([0.296522, -0.671961, -2.814389, -1.226039, 1.570796, 1.867318],accel_mss,speed_ms,0,blend_radius_m)
  movel([0.298113, -0.668161, -2.814797, -1.229430, 1.570796, 1.868909],accel_mss,speed_ms,0,blend_radius_m)
  movel([0.300079, -0.664232, -2.815214, -1.232943, 1.570796, 1.870875],accel_mss,speed_ms,0,blend_radius_m)
  movel([0.301662, -0.661470, -2.815503, -1.235416, 1.570796, 1.872459],accel_mss,speed_ms,0,blend_radius_m)
  movel([0.303456, -0.658709, -2.815788, -1.237892, 1.570796, 1.874252],accel_mss,speed_ms,0,blend_radius_m)
  movel([0.305446, -0.656063, -2.816059, -1.240267, 1.570796, 1.876242],accel_mss,speed_ms,0,blend_radius_m)
  movel([0.307642, -0.653616, -2.816307, -1.242466, 1.570796, 1.878438],accel_mss,speed_ms,0,blend_radius_m)
  movel([0.309571, -0.651910, -2.816478, -1.244001, 1.570796, 1.880367],accel_mss,speed_ms,0,blend_radius_m)
  movel([0.311622, -0.650506, -2.816618, -1.245265, 1.570796, 1.882418],accel_mss,speed_ms,0,blend_radius_m)
  movel([0.313735, -0.649368, -2.816731, -1.246290, 1.570796, 1.884531],accel_mss,speed_ms,0,blend_radius_m)
  movel([0.315866, -0.648458, -2.816821, -1.247110, 1.570796, 1.886662],accel_mss,speed_ms,0,blend_radius_m)
  movel([0.319952, -0.647162, -2.816948, -1.248279, 1.570796, 1.890749],accel_mss,speed_ms,0,blend_radius_m)
  movel([0.323464, -0.646311, -2.817032, -1.249046, 1.570796, 1.894260],accel_mss,speed_ms,0,blend_radius_m)
  movel([0.320966, -0.647160, -2.816948, -1.248281, 1.570796, 1.891763],accel_mss,speed_ms,0,blend_radius_m)
  movel([0.318294, -0.648588, -2.816808, -1.246993, 1.570796, 1.889090],accel_mss,speed_ms,0,blend_radius_m)
  movel([0.315495, -0.650633, -2.816605, -1.245151, 1.570796, 1.886291],accel_mss,speed_ms,0,blend_radius_m)
  movel([0.312607, -0.653345, -2.816334, -1.242710, 1.570796, 1.883404],accel_mss,speed_ms,0,blend_radius_m)
  movel([0.310230, -0.656101, -2.816055, -1.240233, 1.570796, 1.881027],accel_mss,speed_ms,0,blend_radius_m)
  movel([0.308059, -0.659041, -2.815754, -1.237594, 1.570796, 1.878855],accel_mss,speed_ms,0,blend_radius_m)
  movel([0.306173, -0.661908, -2.815457, -1.235023, 1.570796, 1.876970],accel_mss,speed_ms,0,blend_radius_m)
  movel([0.304516, -0.664778, -2.815156, -1.232455, 1.570796, 1.875313],accel_mss,speed_ms,0,blend_radius_m)
  movel([0.301852, -0.670432, -2.814554, -1.227403, 1.570796, 1.872648],accel_mss,speed_ms,0,blend_radius_m)
  movel([0.300013, -0.675802, -2.813969, -1.222618, 1.570796, 1.870810],accel_mss,speed_ms,0,blend_radius_m)
  movel([0.298883, -0.681109, -2.813379, -1.217901, 1.570796, 1.869680],accel_mss,speed_ms,0,blend_radius_m)
  speed_ms = 0.005
  movel([0.298883, -0.674303, -2.806699, -1.231387, 1.570796, 1.869680],accel_mss,speed_ms,0,blend_radius_m)
  speed_ms = 0.040
  movel([0.307826, -0.660581, -2.808192, -1.243616, 1.570796, 1.878622],accel_mss,speed_ms,0,blend_radius_m)
  speed_ms = 0.005
  movel([0.307826, -0.667183, -2.814902, -1.230304, 1.570796, 1.878622],accel_mss,speed_ms,0,blend_radius_m)
  speed_ms = 0.025
  movel([0.307323, -0.668075, -2.814807, -1.229507, 1.570796, 1.878120],accel_mss,speed_ms,0,blend_radius_m)
  movel([0.306534, -0.668662, -2.814744, -1.228983, 1.570796, 1.877330],accel_mss,speed_ms,0,blend_radius_m)
  movel([0.306123, -0.668442, -2.814767, -1.229179, 1.570796, 1.876919],accel_mss,speed_ms,0,blend_radius_m)
  movel([0.306171, -0.667702, -2.814847, -1.229841, 1.570796, 1.876967],accel_mss,speed_ms,0,blend_radius_m)
  movel([0.307220, -0.665774, -2.815051, -1.231564, 1.570796, 1.878017],accel_mss,speed_ms,0,blend_radius_m)
  movel([0.307888, -0.664952, -2.815138, -1.232299, 1.570796, 1.878685],accel_mss,speed_ms,0,blend_radius_m)
  movel([0.308573, -0.664645, -2.815170, -1.232573, 1.570796, 1.879369],accel_mss,speed_ms,0,blend_radius_m)
  movel([0.308862, -0.665041, -2.815129, -1.232219, 1.570796, 1.879658],accel_mss,speed_ms,0,blend_radius_m)
  movel([0.308310, -0.666769, -2.814946, -1.230674, 1.570796, 1.879106],accel_mss,speed_ms,0,blend_radius_m)
  speed_ms = 0.005
  movel([0.308310, -0.660173, -2.808235, -1.243980, 1.570796, 1.879106],accel_mss,speed_ms,0,blend_radius_m)
  speed_ms = 0.040
  movel([0.304559, -0.680779, -2.805966, -1.225644, 1.570796, 1.875355],accel_mss,speed_ms,0,blend_radius_m)
  speed_ms = 0.005
  movel([0.304559, -0.687679, -2.812632, -1.212078, 1.570796, 1.875355],accel_mss,speed_ms,0,blend_radius_m)
  speed_ms = 0.025
  movel([0.307350, -0.684086, -2.813043, -1.215260, 1.570796, 1.878147],accel_mss,speed_ms,0,blend_radius_m)
  movel([0.309763, -0.680457, -2.813452, -1.218480, 1.570796, 1.880560],accel_mss,speed_ms,0,blend_radius_m)
  movel([0.314630, -0.673117, -2.814263, -1.225009, 1.570796, 1.885426],accel_mss,speed_ms,0,blend_radius_m)
  movel([0.318636, -0.668072, -2.814807, -1.229510, 1.570796, 1.889433],accel_mss,speed_ms,0,blend_radius_m)
  movel([0.331896, -0.653061, -2.816363, -1.242965, 1.570796, 1.902692],accel_mss,speed_ms,0,blend_radius_m)
  movel([0.334477, -0.649741, -2.816694, -1.245954, 1.570796, 1.905274],accel_mss,speed_ms,0,blend_radius_m)
  movel([0.335379, -0.648129, -2.816853, -1.247407, 1.570796, 1.906176],accel_mss,speed_ms,0,blend_radius_m)
  movel([0.335707, -0.646781, -2.816986, -1.248622, 1.570796, 1.906504],accel_mss,speed_ms,0,blend_radius_m)
  movel([0.335153, -0.645915, -2.817070, -1.249403, 1.570796, 1.905949],accel_mss,speed_ms,0,blend_radius_m)
  movel([0.333998, -0.645774, -2.817084, -1.249531, 1.570796, 1.904794],accel_mss,speed_ms,0,blend_radius_m)
  movel([0.332045, -0.646011, -2.817061, -1.249317, 1.570796, 1.902842],accel_mss,speed_ms,0,blend_radius_m)
  movel([0.330008, -0.646792, -2.816985, -1.248613, 1.570796, 1.900805],accel_mss,speed_ms,0,blend_radius_m)
  movel([0.327741, -0.648217, -2.816845, -1.247328, 1.570796, 1.898538],accel_mss,speed_ms,0,blend_radius_m)
  movel([0.325107, -0.650377, -2.816631, -1.245382, 1.570796, 1.895903],accel_mss,speed_ms,0,blend_radius_m)
  movel([0.322275, -0.653158, -2.816353, -1.242878, 1.570796, 1.893072],accel_mss,speed_ms,0,blend_radius_m)
  movel([0.319474, -0.656360, -2.816029, -1.240001, 1.570796, 1.890270],accel_mss,speed_ms,0,blend_radius_m)
  movel([0.316738, -0.659850, -2.815671, -1.236868, 1.570796, 1.887534],accel_mss,speed_ms,0,blend_radius_m)
  movel([0.314093, -0.663532, -2.815287, -1.233570, 1.570796, 1.884890],accel_mss,speed_ms,0,blend_radius_m)
  movel([0.309214, -0.670965, -2.814496, -1.226927, 1.570796, 1.880010],accel_mss,speed_ms,0,blend_radius_m)
  movel([0.305058, -0.677762, -2.813753, -1.220874, 1.570796, 1.875854],accel_mss,speed_ms,0,blend_radius_m)
  movel([0.297750, -0.690250, -2.812334, -1.209805, 1.570796, 1.868546],accel_mss,speed_ms,0,blend_radius_m)
  movel([0.295156, -0.694342, -2.811855, -1.206192, 1.570796, 1.865953],accel_mss,speed_ms,0,blend_radius_m)
  movel([0.292310, -0.698383, -2.811374, -1.202631, 1.570796, 1.863107],accel_mss,speed_ms,0,blend_radius_m)
  movel([0.289213, -0.702228, -2.810910, -1.199251, 1.570796, 1.860010],accel_mss,speed_ms,0,blend_radius_m)
  movel([0.285948, -0.705663, -2.810490, -1.196235, 1.570796, 1.856744],accel_mss,speed_ms,0,blend_radius_m)
  movel([0.282594, -0.708480, -2.810142, -1.193767, 1.570796, 1.853391],accel_mss,speed_ms,0,blend_radius_m)
  movel([0.285026, -0.707376, -2.810279, -1.194734, 1.570796, 1.855822],accel_mss,speed_ms,0,blend_radius_m)
  movel([0.287555, -0.705964, -2.810453, -1.195971, 1.570796, 1.858351],accel_mss,speed_ms,0,blend_radius_m)
  movel([0.290159, -0.704250, -2.810664, -1.197475, 1.570796, 1.860956],accel_mss,speed_ms,0,blend_radius_m)
  movel([0.292797, -0.702266, -2.810906, -1.199217, 1.570796, 1.863593],accel_mss,speed_ms,0,blend_radius_m)
  movel([0.292190, -0.705364, -2.810527, -1.196498, 1.570796, 1.862987],accel_mss,speed_ms,0,blend_radius_m)
  movel([0.291131, -0.708713, -2.810113, -1.193562, 1.570796, 1.861928],accel_mss,speed_ms,0,blend_radius_m)
  movel([0.289656, -0.712225, -2.809673, -1.190490, 1.570796, 1.860452],accel_mss,speed_ms,0,blend_radius_m)
  movel([0.287799, -0.715817, -2.809218, -1.187354, 1.570796, 1.858595],accel_mss,speed_ms,0,blend_radius_m)
  movel([0.290896, -0.712003, -2.809701, -1.190684, 1.570796, 1.861693],accel_mss,speed_ms,0,blend_radius_m)
  movel([0.293713, -0.708050, -2.810195, -1.194143, 1.570796, 1.864509],accel_mss,speed_ms,0,blend_radius_m)
  movel([0.296264, -0.703989, -2.810696, -1.197704, 1.570796, 1.867061],accel_mss,speed_ms,0,blend_radius_m)
  movel([0.298581, -0.699851, -2.811198, -1.201340, 1.570796, 1.869377],accel_mss,speed_ms,0,blend_radius_m)
  movel([0.298272, -0.701880, -2.810953, -1.199556, 1.570796, 1.869068],accel_mss,speed_ms,0,blend_radius_m)
  movel([0.297501, -0.704346, -2.810652, -1.197391, 1.570796, 1.868297],accel_mss,speed_ms,0,blend_radius_m)
  movel([0.292554, -0.715994, -2.809195, -1.187199, 1.570796, 1.863350],accel_mss,speed_ms,0,blend_radius_m)
  movel([0.291541, -0.718743, -2.808843, -1.184803, 1.570796, 1.862338],accel_mss,speed_ms,0,blend_radius_m)
  movel([0.290895, -0.721177, -2.808528, -1.182685, 1.570796, 1.861691],accel_mss,speed_ms,0,blend_radius_m)
  movel([0.292970, -0.717075, -2.809057, -1.186257, 1.570796, 1.863766],accel_mss,speed_ms,0,blend_radius_m)
  movel([0.295199, -0.713197, -2.809551, -1.189641, 1.570796, 1.865996],accel_mss,speed_ms,0,blend_radius_m)
  movel([0.300007, -0.705855, -2.810467, -1.196067, 1.570796, 1.870804],accel_mss,speed_ms,0,blend_radius_m)
  movel([0.305109, -0.698569, -2.811352, -1.202467, 1.570796, 1.875905],accel_mss,speed_ms,0,blend_radius_m)
  movel([0.310320, -0.690727, -2.812279, -1.209383, 1.570796, 1.881117],accel_mss,speed_ms,0,blend_radius_m)
  movel([0.313168, -0.685806, -2.812847, -1.213736, 1.570796, 1.883964],accel_mss,speed_ms,0,blend_radius_m)
  movel([0.314986, -0.683051, -2.813160, -1.216178, 1.570796, 1.885783],accel_mss,speed_ms,0,blend_radius_m)
  movel([0.315838, -0.682025, -2.813276, -1.217088, 1.570796, 1.886634],accel_mss,speed_ms,0,blend_radius_m)
  movel([0.316599, -0.681389, -2.813348, -1.217653, 1.570796, 1.887396],accel_mss,speed_ms,0,blend_radius_m)
  movel([0.317214, -0.681212, -2.813367, -1.217809, 1.570796, 1.888010],accel_mss,speed_ms,0,blend_radius_m)
  movel([0.317670, -0.681428, -2.813343, -1.217617, 1.570796, 1.888466],accel_mss,speed_ms,0,blend_radius_m)
  movel([0.318149, -0.682687, -2.813201, -1.216501, 1.570796, 1.888946],accel_mss,speed_ms,0,blend_radius_m)
  movel([0.318083, -0.684506, -2.812995, -1.214888, 1.570796, 1.888880],accel_mss,speed_ms,0,blend_radius_m)
  movel([0.317519, -0.686229, -2.812798, -1.213362, 1.570796, 1.888316],accel_mss,speed_ms,0,blend_radius_m)
  movel([0.320699, -0.680003, -2.813503, -1.218883, 1.570796, 1.891495],accel_mss,speed_ms,0,blend_radius_m)
  movel([0.323397, -0.673856, -2.814182, -1.224350, 1.570796, 1.894193],accel_mss,speed_ms,0,blend_radius_m)
  movel([0.325579, -0.667884, -2.814827, -1.229678, 1.570796, 1.896375],accel_mss,speed_ms,0,blend_radius_m)
  movel([0.327197, -0.662175, -2.815429, -1.234785, 1.570796, 1.897993],accel_mss,speed_ms,0,blend_radius_m)
  speed_ms = 0.005
  movel([0.327197, -0.655648, -2.808710, -1.248031, 1.570796, 1.897993],accel_mss,speed_ms,0,blend_radius_m)
  speed_ms = 0.040
  movel([0.331771, -0.655883, -2.808685, -1.247821, 1.570796, 1.902567],accel_mss,speed_ms,0,blend_radius_m)
  speed_ms = 0.005
  movel([0.331771, -0.662414, -2.815404, -1.234571, 1.570796, 1.902567],accel_mss,speed_ms,0,blend_radius_m)
  speed_ms = 0.025
  movel([0.334530, -0.662229, -2.815424, -1.234736, 1.570796, 1.905327],accel_mss,speed_ms,0,blend_radius_m)
  movel([0.335469, -0.662728, -2.815372, -1.234289, 1.570796, 1.906265],accel_mss,speed_ms,0,blend_radius_m)
  movel([0.335833, -0.663875, -2.815251, -1.233262, 1.570796, 1.906629],accel_mss,speed_ms,0,blend_radius_m)
  movel([0.335591, -0.665349, -2.815096, -1.231944, 1.570796, 1.906388],accel_mss,speed_ms,0,blend_radius_m)
  movel([0.326578, -0.692331, -2.812091, -1.207966, 1.570796, 1.897374],accel_mss,speed_ms,0,blend_radius_m)
  movel([0.325852, -0.694273, -2.811863, -1.206253, 1.570796, 1.896648],accel_mss,speed_ms,0,blend_radius_m)
  movel([0.324885, -0.696285, -2.811625, -1.204479, 1.570796, 1.895681],accel_mss,speed_ms,0,blend_radius_m)
  movel([0.323657, -0.698124, -2.811405, -1.202859, 1.570796, 1.894453],accel_mss,speed_ms,0,blend_radius_m)
  movel([0.322169, -0.699540, -2.811235, -1.201613, 1.570796, 1.892965],accel_mss,speed_ms,0,blend_radius_m)
  movel([0.320845, -0.700147, -2.811162, -1.201079, 1.570796, 1.891642],accel_mss,speed_ms,0,blend_radius_m)
  movel([0.318504, -0.700452, -2.811126, -1.200812, 1.570796, 1.889300],accel_mss,speed_ms,0,blend_radius_m)
  movel([0.317175, -0.701124, -2.811044, -1.200220, 1.570796, 1.887972],accel_mss,speed_ms,0,blend_radius_m)
  movel([0.315504, -0.702819, -2.810839, -1.198732, 1.570796, 1.886301],accel_mss,speed_ms,0,blend_radius_m)
  movel([0.313959, -0.704843, -2.810591, -1.196954, 1.570796, 1.884756],accel_mss,speed_ms,0,blend_radius_m)
  movel([0.312038, -0.707130, -2.810309, -1.194950, 1.570796, 1.882835],accel_mss,speed_ms,0,blend_radius_m)
  movel([0.309999, -0.709150, -2.810059, -1.193180, 1.570796, 1.880795],accel_mss,speed_ms,0,blend_radius_m)
  movel([0.307917, -0.710859, -2.809845, -1.191685, 1.570796, 1.878713],accel_mss,speed_ms,0,blend_radius_m)
  movel([0.305858, -0.712220, -2.809674, -1.190495, 1.570796, 1.876655],accel_mss,speed_ms,0,blend_radius_m)
  movel([0.303892, -0.713197, -2.809551, -1.189642, 1.570796, 1.874689],accel_mss,speed_ms,0,blend_radius_m)
  movel([0.302101, -0.713736, -2.809483, -1.189170, 1.570796, 1.872898],accel_mss,speed_ms,0,blend_radius_m)
  movel([0.300546, -0.713815, -2.809472, -1.189101, 1.570796, 1.871343],accel_mss,speed_ms,0,blend_radius_m)
  movel([0.299304, -0.713373, -2.809528, -1.189487, 1.570796, 1.870100],accel_mss,speed_ms,0,blend_radius_m)
  speed_ms = 0.005
  movel([0.299304, -0.706118, -2.802922, -1.203349, 1.570796, 1.870100],accel_mss,speed_ms,0,blend_radius_m)
  speed_ms = 0.040
  movel([0.281741, -0.732595, -2.799430, -1.180364, 1.570796, 1.852537],accel_mss,speed_ms,0,blend_radius_m)
  speed_ms = 0.005
  movel([0.281741, -0.740198, -2.805971, -1.166219, 1.570796, 1.852537],accel_mss,speed_ms,0,blend_radius_m)
  speed_ms = 0.025
  movel([0.278055, -0.763163, -2.802658, -1.146567, 1.570796, 1.848852],accel_mss,speed_ms,0,blend_radius_m)
  movel([0.277347, -0.766097, -2.802217, -1.144076, 1.570796, 1.848143],accel_mss,speed_ms,0,blend_radius_m)
  movel([0.276648, -0.767628, -2.801985, -1.142777, 1.570796, 1.847444],accel_mss,speed_ms,0,blend_radius_m)
  movel([0.275612, -0.769107, -2.801759, -1.141523, 1.570796, 1.846408],accel_mss,speed_ms,0,blend_radius_m)
  movel([0.272899, -0.771899, -2.801331, -1.139159, 1.570796, 1.843695],accel_mss,speed_ms,0,blend_radius_m)
  movel([0.271996, -0.773553, -2.801075, -1.137761, 1.570796, 1.842792],accel_mss,speed_ms,0,blend_radius_m)
  movel([0.271579, -0.775120, -2.800832, -1.136437, 1.570796, 1.842375],accel_mss,speed_ms,0,blend_radius_m)
  movel([0.271570, -0.777317, -2.800489, -1.134583, 1.570796, 1.842366],accel_mss,speed_ms,0,blend_radius_m)
  movel([0.272150, -0.779102, -2.800208, -1.133079, 1.570796, 1.842946],accel_mss,speed_ms,0,blend_radius_m)
  movel([0.273739, -0.782156, -2.799725, -1.130508, 1.570796, 1.844535],accel_mss,speed_ms,0,blend_radius_m)
  movel([0.274278, -0.784652, -2.799326, -1.128411, 1.570796, 1.845075],accel_mss,speed_ms,0,blend_radius_m)
  movel([0.274468, -0.788653, -2.798680, -1.125056, 1.570796, 1.845264],accel_mss,speed_ms,0,blend_radius_m)
  movel([0.274204, -0.790675, -2.798350, -1.123364, 1.570796, 1.845000],accel_mss,speed_ms,0,blend_radius_m)
  movel([0.273576, -0.792439, -2.798061, -1.121889, 1.570796, 1.844372],accel_mss,speed_ms,0,blend_radius_m)
  movel([0.273096, -0.793150, -2.797944, -1.121295, 1.570796, 1.843892],accel_mss,speed_ms,0,blend_radius_m)
  movel([0.272493, -0.793721, -2.797850, -1.120818, 1.570796, 1.843289],accel_mss,speed_ms,0,blend_radius_m)
  movel([0.271753, -0.794121, -2.797784, -1.120484, 1.570796, 1.842549],accel_mss,speed_ms,0,blend_radius_m)
  movel([0.270866, -0.794320, -2.797751, -1.120318, 1.570796, 1.841663],accel_mss,speed_ms,0,blend_radius_m)
  movel([0.270373, -0.796155, -2.797447, -1.118788, 1.570796, 1.841169],accel_mss,speed_ms,0,blend_radius_m)
  movel([0.270264, -0.798006, -2.797138, -1.117245, 1.570796, 1.841060],accel_mss,speed_ms,0,blend_radius_m)
  movel([0.270864, -0.801605, -2.796533, -1.114251, 1.570796, 1.841661],accel_mss,speed_ms,0,blend_radius_m)
  movel([0.272032, -0.804761, -2.795996, -1.111632, 1.570796, 1.842829],accel_mss,speed_ms,0,blend_radius_m)
  movel([0.273153, -0.807107, -2.795594, -1.109688, 1.570796, 1.843949],accel_mss,speed_ms,0,blend_radius_m)
  movel([0.274846, -0.809256, -2.795223, -1.107909, 1.570796, 1.845642],accel_mss,speed_ms,0,blend_radius_m)
  movel([0.276926, -0.811149, -2.794895, -1.106345, 1.570796, 1.847722],accel_mss,speed_ms,0,blend_radius_m)
  movel([0.278568, -0.813443, -2.794494, -1.104452, 1.570796, 1.849364],accel_mss,speed_ms,0,blend_radius_m)
  movel([0.278969, -0.814935, -2.794232, -1.103222, 1.570796, 1.849766],accel_mss,speed_ms,0,blend_radius_m)
  movel([0.278953, -0.816767, -2.793908, -1.101713, 1.570796, 1.849750],accel_mss,speed_ms,0,blend_radius_m)
  movel([0.278680, -0.817873, -2.793712, -1.100804, 1.570796, 1.849477],accel_mss,speed_ms,0,blend_radius_m)
  movel([0.278145, -0.819070, -2.793499, -1.099820, 1.570796, 1.848941],accel_mss,speed_ms,0,blend_radius_m)
  movel([0.277410, -0.820110, -2.793313, -1.098966, 1.570796, 1.848207],accel_mss,speed_ms,0,blend_radius_m)
  movel([0.276534, -0.820757, -2.793198, -1.098434, 1.570796, 1.847330],accel_mss,speed_ms,0,blend_radius_m)
  movel([0.275921, -0.820812, -2.793188, -1.098389, 1.570796, 1.846718],accel_mss,speed_ms,0,blend_radius_m)
  movel([0.275468, -0.820586, -2.793228, -1.098575, 1.570796, 1.846264],accel_mss,speed_ms,0,blend_radius_m)
  movel([0.271858, -0.817475, -2.793783, -1.101131, 1.570796, 1.842655],accel_mss,speed_ms,0,blend_radius_m)
  movel([0.270330, -0.815583, -2.794118, -1.102688, 1.570796, 1.841127],accel_mss,speed_ms,0,blend_radius_m)
  movel([0.269001, -0.813463, -2.794491, -1.104435, 1.570796, 1.839798],accel_mss,speed_ms,0,blend_radius_m)
  movel([0.268223, -0.814678, -2.794277, -1.103433, 1.570796, 1.839019],accel_mss,speed_ms,0,blend_radius_m)
  movel([0.267662, -0.815894, -2.794063, -1.102432, 1.570796, 1.838458],accel_mss,speed_ms,0,blend_radius_m)
  movel([0.267117, -0.818296, -2.793637, -1.100456, 1.570796, 1.837913],accel_mss,speed_ms,0,blend_radius_m)
  movel([0.267194, -0.820618, -2.793222, -1.098548, 1.570796, 1.837990],accel_mss,speed_ms,0,blend_radius_m)
  movel([0.267740, -0.822801, -2.792830, -1.096758, 1.570796, 1.838537],accel_mss,speed_ms,0,blend_radius_m)
  movel([0.269558, -0.826581, -2.792145, -1.093663, 1.570796, 1.840354],accel_mss,speed_ms,0,blend_radius_m)
  movel([0.271292, -0.829208, -2.791664, -1.091517, 1.570796, 1.842088],accel_mss,speed_ms,0,blend_radius_m)
  movel([0.271782, -0.830334, -2.791456, -1.090598, 1.570796, 1.842578],accel_mss,speed_ms,0,blend_radius_m)
  movel([0.271770, -0.831071, -2.791320, -1.089997, 1.570796, 1.842567],accel_mss,speed_ms,0,blend_radius_m)
  movel([0.271447, -0.831963, -2.791155, -1.089271, 1.570796, 1.842243],accel_mss,speed_ms,0,blend_radius_m)
  movel([0.270811, -0.832930, -2.790976, -1.088483, 1.570796, 1.841608],accel_mss,speed_ms,0,blend_radius_m)
  movel([0.270166, -0.833530, -2.790864, -1.087994, 1.570796, 1.840962],accel_mss,speed_ms,0,blend_radius_m)
  movel([0.268900, -0.834003, -2.790776, -1.087610, 1.570796, 1.839696],accel_mss,speed_ms,0,blend_radius_m)
  movel([0.267192, -0.834426, -2.790697, -1.087266, 1.570796, 1.837988],accel_mss,speed_ms,0,blend_radius_m)
  movel([0.266720, -0.834890, -2.790611, -1.086888, 1.570796, 1.837517],accel_mss,speed_ms,0,blend_radius_m)
  movel([0.266266, -0.835734, -2.790453, -1.086203, 1.570796, 1.837062],accel_mss,speed_ms,0,blend_radius_m)
  movel([0.266043, -0.836616, -2.790287, -1.085486, 1.570796, 1.836840],accel_mss,speed_ms,0,blend_radius_m)
  movel([0.266116, -0.838380, -2.789955, -1.084054, 1.570796, 1.836912],accel_mss,speed_ms,0,blend_radius_m)
  movel([0.266945, -0.841137, -2.789432, -1.081820, 1.570796, 1.837741],accel_mss,speed_ms,0,blend_radius_m)
  movel([0.269138, -0.846567, -2.788390, -1.077432, 1.570796, 1.839934],accel_mss,speed_ms,0,blend_radius_m)
  movel([0.271450, -0.851847, -2.787361, -1.073180, 1.570796, 1.842246],accel_mss,speed_ms,0,blend_radius_m)
  movel([0.271715, -0.853092, -2.787117, -1.072181, 1.570796, 1.842512],accel_mss,speed_ms,0,blend_radius_m)
  movel([0.271667, -0.854575, -2.786823, -1.070990, 1.570796, 1.842463],accel_mss,speed_ms,0,blend_radius_m)
  movel([0.271156, -0.856157, -2.786510, -1.069722, 1.570796, 1.841952],accel_mss,speed_ms,0,blend_radius_m)
  movel([0.270689, -0.856934, -2.786355, -1.069100, 1.570796, 1.841485],accel_mss,speed_ms,0,blend_radius_m)
  movel([0.269378, -0.858253, -2.786092, -1.068044, 1.570796, 1.840175],accel_mss,speed_ms,0,blend_radius_m)
  movel([0.268742, -0.858613, -2.786020, -1.067756, 1.570796, 1.839539],accel_mss,speed_ms,0,blend_radius_m)
  movel([0.267584, -0.858805, -2.785981, -1.067603, 1.570796, 1.838380],accel_mss,speed_ms,0,blend_radius_m)
  movel([0.266607, -0.858483, -2.786046, -1.067860, 1.570796, 1.837403],accel_mss,speed_ms,0,blend_radius_m)
  movel([0.265848, -0.857855, -2.786171, -1.068363, 1.570796, 1.836644],accel_mss,speed_ms,0,blend_radius_m)
  movel([0.262076, -0.853323, -2.787071, -1.071995, 1.570796, 1.832873],accel_mss,speed_ms,0,blend_radius_m)
  movel([0.258644, -0.848379, -2.788039, -1.075971, 1.570796, 1.829441],accel_mss,speed_ms,0,blend_radius_m)
  movel([0.255575, -0.843014, -2.789074, -1.080301, 1.570796, 1.826371],accel_mss,speed_ms,0,blend_radius_m)
  movel([0.252877, -0.837230, -2.790172, -1.084987, 1.570796, 1.823673],accel_mss,speed_ms,0,blend_radius_m)
  movel([0.252039, -0.834921, -2.790605, -1.086863, 1.570796, 1.822835],accel_mss,speed_ms,0,blend_radius_m)
  movel([0.251666, -0.832209, -2.791110, -1.089070, 1.570796, 1.822462],accel_mss,speed_ms,0,blend_radius_m)
  movel([0.251810, -0.830330, -2.791457, -1.090602, 1.570796, 1.822606],accel_mss,speed_ms,0,blend_radius_m)
  movel([0.252185, -0.828305, -2.791830, -1.092255, 1.570796, 1.822981],accel_mss,speed_ms,0,blend_radius_m)
  movel([0.253320, -0.824020, -2.792610, -1.095759, 1.570796, 1.824117],accel_mss,speed_ms,0,blend_radius_m)
  movel([0.258739, -0.807939, -2.795451, -1.108999, 1.570796, 1.829535],accel_mss,speed_ms,0,blend_radius_m)
  movel([0.259950, -0.803494, -2.796212, -1.112683, 1.570796, 1.830746],accel_mss,speed_ms,0,blend_radius_m)
  movel([0.260608, -0.799676, -2.796858, -1.115855, 1.570796, 1.831404],accel_mss,speed_ms,0,blend_radius_m)
  movel([0.260657, -0.798127, -2.797118, -1.117144, 1.570796, 1.831453],accel_mss,speed_ms,0,blend_radius_m)
  movel([0.260469, -0.796893, -2.797324, -1.118172, 1.570796, 1.831265],accel_mss,speed_ms,0,blend_radius_m)
  movel([0.260019, -0.796019, -2.797469, -1.118901, 1.570796, 1.830816],accel_mss,speed_ms,0,blend_radius_m)
  movel([0.259280, -0.795557, -2.797546, -1.119286, 1.570796, 1.830076],accel_mss,speed_ms,0,blend_radius_m)
  movel([0.257564, -0.795430, -2.797567, -1.119392, 1.570796, 1.828361],accel_mss,speed_ms,0,blend_radius_m)
  movel([0.256825, -0.795232, -2.797600, -1.119557, 1.570796, 1.827621],accel_mss,speed_ms,0,blend_radius_m)
  movel([0.256410, -0.794643, -2.797697, -1.120048, 1.570796, 1.827206],accel_mss,speed_ms,0,blend_radius_m)
  movel([0.256635, -0.793038, -2.797963, -1.121389, 1.570796, 1.827431],accel_mss,speed_ms,0,blend_radius_m)
  movel([0.257472, -0.791084, -2.798283, -1.123022, 1.570796, 1.828269],accel_mss,speed_ms,0,blend_radius_m)
  movel([0.260367, -0.784760, -2.799308, -1.128320, 1.570796, 1.831164],accel_mss,speed_ms,0,blend_radius_m)
  movel([0.262974, -0.778509, -2.800302, -1.133578, 1.570796, 1.833770],accel_mss,speed_ms,0,blend_radius_m)
  movel([0.265331, -0.772306, -2.801268, -1.138815, 1.570796, 1.836127],accel_mss,speed_ms,0,blend_radius_m)
  movel([0.267477, -0.766135, -2.802211, -1.144043, 1.570796, 1.838273],accel_mss,speed_ms,0,blend_radius_m)
  movel([0.271335, -0.753816, -2.804037, -1.154536, 1.570796, 1.842131],accel_mss,speed_ms,0,blend_radius_m)
  movel([0.274904, -0.741375, -2.805808, -1.165206, 1.570796, 1.845701],accel_mss,speed_ms,0,blend_radius_m)
  speed_ms = 0.005
  movel([0.274904, -0.733757, -2.799270, -1.179362, 1.570796, 1.845701],accel_mss,speed_ms,0,blend_radius_m)
  speed_ms = 0.040
  movel([0.261432, -0.765815, -2.794583, -1.151992, 1.570796, 1.832228],accel_mss,speed_ms,0,blend_radius_m)
  speed_ms = 0.005
  movel([0.261432, -0.773820, -2.801034, -1.137534, 1.570796, 1.832228],accel_mss,speed_ms,0,blend_radius_m)
  speed_ms = 0.025
  movel([0.254948, -0.782417, -2.799683, -1.130289, 1.570796, 1.825745],accel_mss,speed_ms,0,blend_radius_m)
  movel([0.248348, -0.790765, -2.798335, -1.123288, 1.570796, 1.819145],accel_mss,speed_ms,0,blend_radius_m)
  movel([0.241644, -0.798860, -2.796995, -1.116534, 1.570796, 1.812440],accel_mss,speed_ms,0,blend_radius_m)
  movel([0.234856, -0.806677, -2.795668, -1.110044, 1.570796, 1.805652],accel_mss,speed_ms,0,blend_radius_m)
  movel([0.240164, -0.798666, -2.797027, -1.116696, 1.570796, 1.810961],accel_mss,speed_ms,0,blend_radius_m)
  movel([0.245154, -0.790478, -2.798382, -1.123529, 1.570796, 1.815950],accel_mss,speed_ms,0,blend_radius_m)
  movel([0.249787, -0.782167, -2.799723, -1.130500, 1.570796, 1.820583],accel_mss,speed_ms,0,blend_radius_m)
  movel([0.254028, -0.773788, -2.801039, -1.137562, 1.570796, 1.824825],accel_mss,speed_ms,0,blend_radius_m)
  movel([0.248584, -0.780848, -2.799932, -1.131608, 1.570796, 1.819380],accel_mss,speed_ms,0,blend_radius_m)
  movel([0.243053, -0.787719, -2.798831, -1.125839, 1.570796, 1.813849],accel_mss,speed_ms,0,blend_radius_m)
  movel([0.237436, -0.794399, -2.797738, -1.120252, 1.570796, 1.808232],accel_mss,speed_ms,0,blend_radius_m)
  movel([0.231748, -0.800868, -2.796657, -1.114864, 1.570796, 1.802544],accel_mss,speed_ms,0,blend_radius_m)
  movel([0.225400, -0.807899, -2.795458, -1.109032, 1.570796, 1.796196],accel_mss,speed_ms,0,blend_radius_m)
  movel([0.219321, -0.815081, -2.794206, -1.103102, 1.570796, 1.790117],accel_mss,speed_ms,0,blend_radius_m)
  movel([0.216506, -0.818848, -2.793539, -1.100002, 1.570796, 1.787302],accel_mss,speed_ms,0,blend_radius_m)
  movel([0.213960, -0.822707, -2.792847, -1.096835, 1.570796, 1.784756],accel_mss,speed_ms,0,blend_radius_m)
  movel([0.211819, -0.826568, -2.792147, -1.093674, 1.570796, 1.782615],accel_mss,speed_ms,0,blend_radius_m)
  movel([0.210196, -0.830343, -2.791455, -1.090591, 1.570796, 1.780992],accel_mss,speed_ms,0,blend_radius_m)
  movel([0.211400, -0.825947, -2.792260, -1.094182, 1.570796, 1.782197],accel_mss,speed_ms,0,blend_radius_m)
  movel([0.212956, -0.821288, -2.793102, -1.097999, 1.570796, 1.783752],accel_mss,speed_ms,0,blend_radius_m)
  movel([0.214839, -0.816424, -2.793969, -1.101996, 1.570796, 1.785635],accel_mss,speed_ms,0,blend_radius_m)
  movel([0.217020, -0.811415, -2.794849, -1.106126, 1.570796, 1.787816],accel_mss,speed_ms,0,blend_radius_m)
  movel([0.219468, -0.806323, -2.795729, -1.110337, 1.570796, 1.790265],accel_mss,speed_ms,0,blend_radius_m)
  movel([0.222158, -0.801210, -2.796599, -1.114580, 1.570796, 1.792954],accel_mss,speed_ms,0,blend_radius_m)
  movel([0.225056, -0.796142, -2.797449, -1.118798, 1.570796, 1.795852],accel_mss,speed_ms,0,blend_radius_m)
  movel([0.228128, -0.791192, -2.798266, -1.122931, 1.570796, 1.798924],accel_mss,speed_ms,0,blend_radius_m)
  movel([0.222602, -0.798941, -2.796981, -1.116467, 1.570796, 1.793398],accel_mss,speed_ms,0,blend_radius_m)
  movel([0.217407, -0.806697, -2.795665, -1.110027, 1.570796, 1.788203],accel_mss,speed_ms,0,blend_radius_m)
  movel([0.212522, -0.814438, -2.794319, -1.103632, 1.570796, 1.783318],accel_mss,speed_ms,0,blend_radius_m)
  movel([0.207928, -0.822138, -2.792950, -1.097301, 1.570796, 1.778724],accel_mss,speed_ms,0,blend_radius_m)
  movel([0.203609, -0.829770, -2.791560, -1.091059, 1.570796, 1.774406],accel_mss,speed_ms,0,blend_radius_m)
  movel([0.199541, -0.837315, -2.790156, -1.084918, 1.570796, 1.770338],accel_mss,speed_ms,0,blend_radius_m)
  movel([0.192077, -0.852055, -2.787321, -1.073013, 1.570796, 1.762873],accel_mss,speed_ms,0,blend_radius_m)
  movel([0.194129, -0.847076, -2.788292, -1.077021, 1.570796, 1.764926],accel_mss,speed_ms,0,blend_radius_m)
  movel([0.195772, -0.841860, -2.789294, -1.081234, 1.570796, 1.766568],accel_mss,speed_ms,0,blend_radius_m)
  movel([0.198677, -0.831730, -2.791198, -1.089460, 1.570796, 1.769474],accel_mss,speed_ms,0,blend_radius_m)
  movel([0.200321, -0.827105, -2.792049, -1.093235, 1.570796, 1.771117],accel_mss,speed_ms,0,blend_radius_m)
  movel([0.202086, -0.822857, -2.792820, -1.096712, 1.570796, 1.772882],accel_mss,speed_ms,0,blend_radius_m)
  movel([0.206386, -0.813912, -2.794412, -1.104065, 1.570796, 1.777183],accel_mss,speed_ms,0,blend_radius_m)
  movel([0.205471, -0.815219, -2.794182, -1.102988, 1.570796, 1.776267],accel_mss,speed_ms,0,blend_radius_m)
  movel([0.203922, -0.816927, -2.793880, -1.101582, 1.570796, 1.774718],accel_mss,speed_ms,0,blend_radius_m)
  movel([0.195262, -0.825147, -2.792406, -1.094836, 1.570796, 1.766058],accel_mss,speed_ms,0,blend_radius_m)
  movel([0.192150, -0.828269, -2.791836, -1.092284, 1.570796, 1.762947],accel_mss,speed_ms,0,blend_radius_m)
  movel([0.188692, -0.832669, -2.791024, -1.088696, 1.570796, 1.759489],accel_mss,speed_ms,0,blend_radius_m)
  movel([0.185491, -0.837327, -2.790153, -1.084908, 1.570796, 1.756287],accel_mss,speed_ms,0,blend_radius_m)
  movel([0.179730, -0.846690, -2.788367, -1.077333, 1.570796, 1.750526],accel_mss,speed_ms,0,blend_radius_m)
  movel([0.181985, -0.841843, -2.789298, -1.081248, 1.570796, 1.752782],accel_mss,speed_ms,0,blend_radius_m)
  movel([0.183935, -0.837015, -2.790212, -1.085162, 1.570796, 1.754732],accel_mss,speed_ms,0,blend_radius_m)
  movel([0.187766, -0.827282, -2.792017, -1.093091, 1.570796, 1.758562],accel_mss,speed_ms,0,blend_radius_m)
  movel([0.190156, -0.822112, -2.792954, -1.097322, 1.570796, 1.760953],accel_mss,speed_ms,0,blend_radius_m)
  movel([0.192896, -0.816834, -2.793897, -1.101658, 1.570796, 1.763693],accel_mss,speed_ms,0,blend_radius_m)
  movel([0.199179, -0.806010, -2.795783, -1.110597, 1.570796, 1.769975],accel_mss,speed_ms,0,blend_radius_m)
  movel([0.212906, -0.784126, -2.799410, -1.128853, 1.570796, 1.783702],accel_mss,speed_ms,0,blend_radius_m)
  movel([0.207618, -0.788594, -2.798689, -1.125106, 1.570796, 1.778414],accel_mss,speed_ms,0,blend_radius_m)
  movel([0.202419, -0.793369, -2.797908, -1.121112, 1.570796, 1.773215],accel_mss,speed_ms,0,blend_radius_m)
  movel([0.197333, -0.798410, -2.797070, -1.116909, 1.570796, 1.768130],accel_mss,speed_ms,0,blend_radius_m)
  movel([0.192402, -0.803673, -2.796182, -1.112534, 1.570796, 1.763198],accel_mss,speed_ms,0,blend_radius_m)
  movel([0.187658, -0.809120, -2.795247, -1.108022, 1.570796, 1.758454],accel_mss,speed_ms,0,blend_radius_m)
  movel([0.183125, -0.814720, -2.794270, -1.103399, 1.570796, 1.753921],accel_mss,speed_ms,0,blend_radius_m)
  movel([0.178832, -0.820428, -2.793256, -1.098704, 1.570796, 1.749628],accel_mss,speed_ms,0,blend_radius_m)
  movel([0.174808, -0.826215, -2.792211, -1.093962, 1.570796, 1.745604],accel_mss,speed_ms,0,blend_radius_m)
  movel([0.175871, -0.824454, -2.792531, -1.095404, 1.570796, 1.746668],accel_mss,speed_ms,0,blend_radius_m)
  movel([0.176866, -0.822501, -2.792884, -1.097003, 1.570796, 1.747662],accel_mss,speed_ms,0,blend_radius_m)
  movel([0.178700, -0.818256, -2.793644, -1.100489, 1.570796, 1.749496],accel_mss,speed_ms,0,blend_radius_m)
  movel([0.182052, -0.810100, -2.795077, -1.107212, 1.570796, 1.752849],accel_mss,speed_ms,0,blend_radius_m)
  movel([0.185570, -0.802963, -2.796302, -1.113123, 1.570796, 1.756367],accel_mss,speed_ms,0,blend_radius_m)
  movel([0.189353, -0.795776, -2.797510, -1.119103, 1.570796, 1.760150],accel_mss,speed_ms,0,blend_radius_m)
  movel([0.193392, -0.788541, -2.798698, -1.125150, 1.570796, 1.764188],accel_mss,speed_ms,0,blend_radius_m)
  movel([0.197671, -0.781258, -2.799867, -1.131263, 1.570796, 1.768468],accel_mss,speed_ms,0,blend_radius_m)
  movel([0.202185, -0.773917, -2.801019, -1.137453, 1.570796, 1.772981],accel_mss,speed_ms,0,blend_radius_m)
  movel([0.206927, -0.766523, -2.802152, -1.143714, 1.570796, 1.777723],accel_mss,speed_ms,0,blend_radius_m)
  movel([0.217047, -0.751540, -2.804366, -1.156482, 1.570796, 1.787844],accel_mss,speed_ms,0,blend_radius_m)
  movel([0.212834, -0.756242, -2.803683, -1.152464, 1.570796, 1.783630],accel_mss,speed_ms,0,blend_radius_m)
  movel([0.199928, -0.769519, -2.801696, -1.141174, 1.570796, 1.770724],accel_mss,speed_ms,0,blend_radius_m)
  movel([0.195714, -0.774033, -2.801001, -1.137355, 1.570796, 1.766510],accel_mss,speed_ms,0,blend_radius_m)
  movel([0.191666, -0.778730, -2.800267, -1.133392, 1.570796, 1.762463],accel_mss,speed_ms,0,blend_radius_m)
  movel([0.187933, -0.783588, -2.799496, -1.129305, 1.570796, 1.758729],accel_mss,speed_ms,0,blend_radius_m)
  movel([0.184647, -0.788604, -2.798688, -1.125097, 1.570796, 1.755443],accel_mss,speed_ms,0,blend_radius_m)
  movel([0.189107, -0.780379, -2.800007, -1.132003, 1.570796, 1.759904],accel_mss,speed_ms,0,blend_radius_m)
  movel([0.193566, -0.771802, -2.801346, -1.139241, 1.570796, 1.764363],accel_mss,speed_ms,0,blend_radius_m)
  movel([0.198297, -0.763170, -2.802657, -1.146562, 1.570796, 1.769093],accel_mss,speed_ms,0,blend_radius_m)
  movel([0.200846, -0.758938, -2.803287, -1.150164, 1.570796, 1.771643],accel_mss,speed_ms,0,blend_radius_m)
  movel([0.203569, -0.754815, -2.803892, -1.153682, 1.570796, 1.774365],accel_mss,speed_ms,0,blend_radius_m)
  movel([0.213662, -0.740926, -2.805870, -1.165593, 1.570796, 1.784458],accel_mss,speed_ms,0,blend_radius_m)
  movel([0.224121, -0.726878, -2.807779, -1.177732, 1.570796, 1.794917],accel_mss,speed_ms,0,blend_radius_m)
  movel([0.216555, -0.734218, -2.806793, -1.171378, 1.570796, 1.787351],accel_mss,speed_ms,0,blend_radius_m)
  movel([0.209738, -0.741508, -2.805789, -1.165092, 1.570796, 1.780535],accel_mss,speed_ms,0,blend_radius_m)
  movel([0.203245, -0.749235, -2.804698, -1.158456, 1.570796, 1.774041],accel_mss,speed_ms,0,blend_radius_m)
  movel([0.196669, -0.757856, -2.803446, -1.151087, 1.570796, 1.767465],accel_mss,speed_ms,0,blend_radius_m)
  movel([0.199815, -0.753266, -2.804117, -1.155006, 1.570796, 1.770611],accel_mss,speed_ms,0,blend_radius_m)
  movel([0.202657, -0.748603, -2.804788, -1.158998, 1.570796, 1.773453],accel_mss,speed_ms,0,blend_radius_m)
  movel([0.213090, -0.729443, -2.807437, -1.175509, 1.570796, 1.783886],accel_mss,speed_ms,0,blend_radius_m)
  movel([0.215992, -0.724580, -2.808082, -1.179726, 1.570796, 1.786788],accel_mss,speed_ms,0,blend_radius_m)
  movel([0.219234, -0.719707, -2.808718, -1.183963, 1.570796, 1.790031],accel_mss,speed_ms,0,blend_radius_m)
  movel([0.223935, -0.713458, -2.809518, -1.189413, 1.570796, 1.794731],accel_mss,speed_ms,0,blend_radius_m)
  movel([0.228034, -0.708871, -2.810093, -1.193425, 1.570796, 1.798830],accel_mss,speed_ms,0,blend_radius_m)
  movel([0.228958, -0.707578, -2.810254, -1.194557, 1.570796, 1.799754],accel_mss,speed_ms,0,blend_radius_m)
  movel([0.229281, -0.706484, -2.810389, -1.195516, 1.570796, 1.800078],accel_mss,speed_ms,0,blend_radius_m)
  movel([0.228746, -0.706255, -2.810417, -1.195716, 1.570796, 1.799542],accel_mss,speed_ms,0,blend_radius_m)
  movel([0.227577, -0.706693, -2.810363, -1.195333, 1.570796, 1.798373],accel_mss,speed_ms,0,blend_radius_m)
  movel([0.226000, -0.707607, -2.810250, -1.194532, 1.570796, 1.796796],accel_mss,speed_ms,0,blend_radius_m)
  movel([0.222512, -0.710046, -2.809947, -1.192396, 1.570796, 1.793308],accel_mss,speed_ms,0,blend_radius_m)
  movel([0.220069, -0.711994, -2.809703, -1.190693, 1.570796, 1.790865],accel_mss,speed_ms,0,blend_radius_m)
  movel([0.223947, -0.706331, -2.810408, -1.195650, 1.570796, 1.794743],accel_mss,speed_ms,0,blend_radius_m)
  movel([0.228482, -0.700617, -2.811106, -1.200666, 1.570796, 1.799278],accel_mss,speed_ms,0,blend_radius_m)
  movel([0.237978, -0.689792, -2.812388, -1.210209, 1.570796, 1.808774],accel_mss,speed_ms,0,blend_radius_m)
  speed_ms = 0.005
  movel([0.237978, -0.682863, -2.805726, -1.223800, 1.570796, 1.808774],accel_mss,speed_ms,0,blend_radius_m)
  speed_ms = 0.040
  movel([0.220547, -0.693122, -2.804519, -1.214749, 1.570796, 1.791343],accel_mss,speed_ms,0,blend_radius_m)
  speed_ms = 0.005
  movel([0.220547, -0.700197, -2.811156, -1.201035, 1.570796, 1.791343],accel_mss,speed_ms,0,blend_radius_m)
  speed_ms = 0.025
  movel([0.219117, -0.698802, -2.811324, -1.202263, 1.570796, 1.789913],accel_mss,speed_ms,0,blend_radius_m)
  movel([0.217209, -0.698130, -2.811405, -1.202854, 1.570796, 1.788005],accel_mss,speed_ms,0,blend_radius_m)
  movel([0.214903, -0.698104, -2.811408, -1.202877, 1.570796, 1.785699],accel_mss,speed_ms,0,blend_radius_m)
  movel([0.212279, -0.698634, -2.811344, -1.202411, 1.570796, 1.783076],accel_mss,speed_ms,0,blend_radius_m)
  movel([0.209410, -0.699653, -2.811222, -1.201514, 1.570796, 1.780207],accel_mss,speed_ms,0,blend_radius_m)
  movel([0.206382, -0.701071, -2.811051, -1.200267, 1.570796, 1.777179],accel_mss,speed_ms,0,blend_radius_m)
  movel([0.200145, -0.704773, -2.810600, -1.197016, 1.570796, 1.770941],accel_mss,speed_ms,0,blend_radius_m)
  speed_ms = 0.005
  movel([0.200145, -0.697634, -2.803973, -1.210782, 1.570796, 1.770941],accel_mss,speed_ms,0,blend_radius_m)
  speed_ms = 0.040
  movel([0.225931, -0.675461, -2.806569, -1.230358, 1.570796, 1.796727],accel_mss,speed_ms,0,blend_radius_m)
  speed_ms = 0.005
  movel([0.225931, -0.682284, -2.813247, -1.216858, 1.570796, 1.796727],accel_mss,speed_ms,0,blend_radius_m)
  speed_ms = 0.025
  movel([0.225055, -0.678580, -2.813662, -1.220148, 1.570796, 1.795851],accel_mss,speed_ms,0,blend_radius_m)
  movel([0.223901, -0.675290, -2.814025, -1.223074, 1.570796, 1.794697],accel_mss,speed_ms,0,blend_radius_m)
  movel([0.222358, -0.672573, -2.814322, -1.225494, 1.570796, 1.793155],accel_mss,speed_ms,0,blend_radius_m)
  movel([0.220313, -0.670581, -2.814538, -1.227270, 1.570796, 1.791109],accel_mss,speed_ms,0,blend_radius_m)
  movel([0.217651, -0.669491, -2.814655, -1.228243, 1.570796, 1.788447],accel_mss,speed_ms,0,blend_radius_m)
  movel([0.214276, -0.669435, -2.814661, -1.228292, 1.570796, 1.785072],accel_mss,speed_ms,0,blend_radius_m)
  movel([0.210076, -0.670590, -2.814537, -1.227262, 1.570796, 1.780872],accel_mss,speed_ms,0,blend_radius_m)
  movel([0.207638, -0.671663, -2.814421, -1.226305, 1.570796, 1.778434],accel_mss,speed_ms,0,blend_radius_m)
  movel([0.204957, -0.673094, -2.814266, -1.225030, 1.570796, 1.775753],accel_mss,speed_ms,0,blend_radius_m)
  speed_ms = 0.005
  movel([0.204957, -0.666405, -2.807568, -1.238416, 1.570796, 1.775753],accel_mss,speed_ms,0,blend_radius_m)
  speed_ms = 0.040
  movel([0.226788, -0.648320, -2.809459, -1.254610, 1.570796, 1.797585],accel_mss,speed_ms,0,blend_radius_m)
  speed_ms = 0.005
  movel([0.226788, -0.654735, -2.816194, -1.241461, 1.570796, 1.797585],accel_mss,speed_ms,0,blend_radius_m)
  speed_ms = 0.025
  movel([0.226566, -0.645840, -2.817077, -1.249471, 1.570796, 1.797362],accel_mss,speed_ms,0,blend_radius_m)
  movel([0.225962, -0.641939, -2.817455, -1.252995, 1.570796, 1.796758],accel_mss,speed_ms,0,blend_radius_m)
  movel([0.224859, -0.638608, -2.817772, -1.256009, 1.570796, 1.795656],accel_mss,speed_ms,0,blend_radius_m)
  movel([0.223137, -0.636010, -2.818017, -1.258363, 1.570796, 1.793933],accel_mss,speed_ms,0,blend_radius_m)
  movel([0.220667, -0.634310, -2.818175, -1.259904, 1.570796, 1.791464],accel_mss,speed_ms,0,blend_radius_m)
  movel([0.217324, -0.633662, -2.818235, -1.260492, 1.570796, 1.788120],accel_mss,speed_ms,0,blend_radius_m)
  movel([0.212992, -0.634231, -2.818182, -1.259976, 1.570796, 1.783788],accel_mss,speed_ms,0,blend_radius_m)
  speed_ms = 0.005
  movel([0.212992, -0.628135, -2.811409, -1.272846, 1.570796, 1.783788],accel_mss,speed_ms,0,blend_radius_m)
  speed_ms = 0.040
  movel([0.232327, -0.619609, -2.812182, -1.280598, 1.570796, 1.803124],accel_mss,speed_ms,0,blend_radius_m)
  speed_ms = 0.005
  movel([0.232327, -0.625567, -2.818972, -1.267851, 1.570796, 1.803124],accel_mss,speed_ms,0,blend_radius_m)
  speed_ms = 0.025
  movel([0.233592, -0.619247, -2.819528, -1.273614, 1.570796, 1.804388],accel_mss,speed_ms,0,blend_radius_m)
  movel([0.234489, -0.613055, -2.820058, -1.279275, 1.570796, 1.805285],accel_mss,speed_ms,0,blend_radius_m)
  movel([0.234865, -0.607220, -2.820544, -1.284624, 1.570796, 1.805662],accel_mss,speed_ms,0,blend_radius_m)
  movel([0.234575, -0.601989, -2.820969, -1.289432, 1.570796, 1.805371],accel_mss,speed_ms,0,blend_radius_m)
  movel([0.233465, -0.597590, -2.821317, -1.293482, 1.570796, 1.804261],accel_mss,speed_ms,0,blend_radius_m)
  movel([0.232550, -0.595788, -2.821458, -1.295143, 1.570796, 1.803347],accel_mss,speed_ms,0,blend_radius_m)
  movel([0.229927, -0.593110, -2.821664, -1.297614, 1.570796, 1.800723],accel_mss,speed_ms,0,blend_radius_m)
  movel([0.228177, -0.592302, -2.821726, -1.298361, 1.570796, 1.798973],accel_mss,speed_ms,0,blend_radius_m)
  movel([0.226109, -0.591884, -2.821758, -1.298747, 1.570796, 1.796905],accel_mss,speed_ms,0,blend_radius_m)
  movel([0.223710, -0.591892, -2.821758, -1.298740, 1.570796, 1.794507],accel_mss,speed_ms,0,blend_radius_m)
  speed_ms = 0.005
  movel([0.223710, -0.586490, -2.814912, -1.310987, 1.570796, 1.794507],accel_mss,speed_ms,0,blend_radius_m)
  speed_ms = 0.040
  movel([0.244747, -0.576105, -2.815680, -1.320604, 1.570796, 1.815543],accel_mss,speed_ms,0,blend_radius_m)
  speed_ms = 0.005
  movel([0.244747, -0.581326, -2.822541, -1.308521, 1.570796, 1.815543],accel_mss,speed_ms,0,blend_radius_m)
  speed_ms = 0.025
  movel([0.246755, -0.573573, -2.823090, -1.315727, 1.570796, 1.817551],accel_mss,speed_ms,0,blend_radius_m)
  movel([0.248116, -0.566150, -2.823593, -1.322646, 1.570796, 1.818913],accel_mss,speed_ms,0,blend_radius_m)
  movel([0.248691, -0.559316, -2.824039, -1.329034, 1.570796, 1.819487],accel_mss,speed_ms,0,blend_radius_m)
  movel([0.248301, -0.553370, -2.824413, -1.334606, 1.570796, 1.819097],accel_mss,speed_ms,0,blend_radius_m)
  movel([0.246800, -0.548584, -2.824704, -1.339101, 1.570796, 1.817596],accel_mss,speed_ms,0,blend_radius_m)
  movel([0.245573, -0.546724, -2.824815, -1.340850, 1.570796, 1.816369],accel_mss,speed_ms,0,blend_radius_m)
  movel([0.244017, -0.545253, -2.824902, -1.342234, 1.570796, 1.814813],accel_mss,speed_ms,0,blend_radius_m)
  movel([0.242096, -0.544228, -2.824962, -1.343199, 1.570796, 1.812893],accel_mss,speed_ms,0,blend_radius_m)
  movel([0.239802, -0.543663, -2.824995, -1.343731, 1.570796, 1.810599],accel_mss,speed_ms,0,blend_radius_m)
  movel([0.237118, -0.543609, -2.824998, -1.343782, 1.570796, 1.807915],accel_mss,speed_ms,0,blend_radius_m)
  movel([0.234025, -0.544086, -2.824970, -1.343333, 1.570796, 1.804821],accel_mss,speed_ms,0,blend_radius_m)
  speed_ms = 0.005
  movel([0.234025, -0.539523, -2.818059, -1.354807, 1.570796, 1.804821],accel_mss,speed_ms,0,blend_radius_m)
  speed_ms = 0.040
  movel([0.134268, -0.609479, -2.813063, -1.289847, 1.570796, 1.705065],accel_mss,speed_ms,0,blend_radius_m)
  speed_ms = 0.005
  movel([0.134268, -0.615270, -2.819871, -1.277248, 1.570796, 1.705065],accel_mss,speed_ms,0,blend_radius_m)
  speed_ms = 0.025
  movel([0.139062, -0.615079, -2.819887, -1.277423, 1.570796, 1.709858],accel_mss,speed_ms,0,blend_radius_m)
  movel([0.143343, -0.615724, -2.819832, -1.276833, 1.570796, 1.714139],accel_mss,speed_ms,0,blend_radius_m)
  movel([0.147131, -0.617145, -2.819710, -1.275534, 1.570796, 1.717927],accel_mss,speed_ms,0,blend_radius_m)
  movel([0.150438, -0.619282, -2.819525, -1.273582, 1.570796, 1.721234],accel_mss,speed_ms,0,blend_radius_m)
  movel([0.153266, -0.622083, -2.819280, -1.271026, 1.570796, 1.724062],accel_mss,speed_ms,0,blend_radius_m)
  movel([0.155649, -0.625476, -2.818980, -1.267933, 1.570796, 1.726445],accel_mss,speed_ms,0,blend_radius_m)
  movel([0.157585, -0.629417, -2.818625, -1.264348, 1.570796, 1.728381],accel_mss,speed_ms,0,blend_radius_m)
  movel([0.159113, -0.633822, -2.818220, -1.260347, 1.570796, 1.729909],accel_mss,speed_ms,0,blend_radius_m)
  movel([0.160234, -0.638644, -2.817769, -1.255976, 1.570796, 1.731031],accel_mss,speed_ms,0,blend_radius_m)
  movel([0.160985, -0.643813, -2.817274, -1.251302, 1.570796, 1.731782],accel_mss,speed_ms,0,blend_radius_m)
  movel([0.161377, -0.649266, -2.816741, -1.246382, 1.570796, 1.732173],accel_mss,speed_ms,0,blend_radius_m)
  movel([0.161433, -0.654953, -2.816172, -1.241264, 1.570796, 1.732229],accel_mss,speed_ms,0,blend_radius_m)
  movel([0.161176, -0.660797, -2.815573, -1.236020, 1.570796, 1.731972],accel_mss,speed_ms,0,blend_radius_m)
  movel([0.160617, -0.666761, -2.814947, -1.230682, 1.570796, 1.731414],accel_mss,speed_ms,0,blend_radius_m)
  movel([0.159785, -0.672766, -2.814301, -1.225322, 1.570796, 1.730581],accel_mss,speed_ms,0,blend_radius_m)
  movel([0.158700, -0.678768, -2.813641, -1.219980, 1.570796, 1.729497],accel_mss,speed_ms,0,blend_radius_m)
  movel([0.156908, -0.686907, -2.812721, -1.212761, 1.570796, 1.727704],accel_mss,speed_ms,0,blend_radius_m)
  movel([0.154407, -0.696429, -2.811608, -1.204352, 1.570796, 1.725204],accel_mss,speed_ms,0,blend_radius_m)
  movel([0.151119, -0.706637, -2.810370, -1.195381, 1.570796, 1.721915],accel_mss,speed_ms,0,blend_radius_m)
  movel([0.149156, -0.711788, -2.809728, -1.190873, 1.570796, 1.719952],accel_mss,speed_ms,0,blend_radius_m)
  movel([0.146975, -0.716847, -2.809086, -1.186455, 1.570796, 1.717771],accel_mss,speed_ms,0,blend_radius_m)
  movel([0.144549, -0.721757, -2.808452, -1.182180, 1.570796, 1.715345],accel_mss,speed_ms,0,blend_radius_m)
  movel([0.141880, -0.726416, -2.807840, -1.178133, 1.570796, 1.712676],accel_mss,speed_ms,0,blend_radius_m)
  movel([0.138944, -0.730766, -2.807260, -1.174363, 1.570796, 1.709741],accel_mss,speed_ms,0,blend_radius_m)
  movel([0.135729, -0.734733, -2.806723, -1.170933, 1.570796, 1.706525],accel_mss,speed_ms,0,blend_radius_m)
  movel([0.132223, -0.738233, -2.806243, -1.167913, 1.570796, 1.703020],accel_mss,speed_ms,0,blend_radius_m)
  movel([0.128404, -0.741211, -2.805830, -1.165348, 1.570796, 1.699201],accel_mss,speed_ms,0,blend_radius_m)
  movel([0.126366, -0.742481, -2.805653, -1.164254, 1.570796, 1.697163],accel_mss,speed_ms,0,blend_radius_m)
  movel([0.124243, -0.743598, -2.805497, -1.163295, 1.570796, 1.695039],accel_mss,speed_ms,0,blend_radius_m)
  movel([0.119724, -0.745330, -2.805253, -1.161807, 1.570796, 1.690521],accel_mss,speed_ms,0,blend_radius_m)
  movel([0.114551, -0.746579, -2.805076, -1.160734, 1.570796, 1.685347],accel_mss,speed_ms,0,blend_radius_m)
  movel([0.109817, -0.747182, -2.804990, -1.160217, 1.570796, 1.680614],accel_mss,speed_ms,0,blend_radius_m)
  movel([0.105467, -0.747216, -2.804985, -1.160188, 1.570796, 1.676263],accel_mss,speed_ms,0,blend_radius_m)
  movel([0.101426, -0.746746, -2.805052, -1.160591, 1.570796, 1.672223],accel_mss,speed_ms,0,blend_radius_m)
  movel([0.097644, -0.745837, -2.805181, -1.161371, 1.570796, 1.668440],accel_mss,speed_ms,0,blend_radius_m)
  movel([0.094051, -0.744565, -2.805361, -1.162463, 1.570796, 1.664847],accel_mss,speed_ms,0,blend_radius_m)
  movel([0.087186, -0.741198, -2.805832, -1.165359, 1.570796, 1.657982],accel_mss,speed_ms,0,blend_radius_m)
  movel([0.079841, -0.737147, -2.806393, -1.168849, 1.570796, 1.650638],accel_mss,speed_ms,0,blend_radius_m)
  movel([0.072694, -0.732912, -2.806970, -1.172507, 1.570796, 1.643490],accel_mss,speed_ms,0,blend_radius_m)
  movel([0.065973, -0.728094, -2.807617, -1.176678, 1.570796, 1.636769],accel_mss,speed_ms,0,blend_radius_m)
  movel([0.062851, -0.725329, -2.807984, -1.179077, 1.570796, 1.633647],accel_mss,speed_ms,0,blend_radius_m)
  movel([0.059928, -0.722251, -2.808388, -1.181750, 1.570796, 1.630725],accel_mss,speed_ms,0,blend_radius_m)
  movel([0.056167, -0.718564, -2.808866, -1.184960, 1.570796, 1.626963],accel_mss,speed_ms,0,blend_radius_m)
  movel([0.051841, -0.715427, -2.809268, -1.187694, 1.570796, 1.622637],accel_mss,speed_ms,0,blend_radius_m)
  movel([0.047031, -0.712809, -2.809600, -1.189980, 1.570796, 1.617827],accel_mss,speed_ms,0,blend_radius_m)
  movel([0.041837, -0.710642, -2.809872, -1.191875, 1.570796, 1.612633],accel_mss,speed_ms,0,blend_radius_m)
  movel([0.030653, -0.707469, -2.810267, -1.194652, 1.570796, 1.601450],accel_mss,speed_ms,0,blend_radius_m)
  movel([0.019045, -0.705425, -2.810520, -1.196445, 1.570796, 1.589842],accel_mss,speed_ms,0,blend_radius_m)
  movel([0.009832, -0.704717, -2.810607, -1.197065, 1.570796, 1.580628],accel_mss,speed_ms,0,blend_radius_m)
  movel([-0.000049, -0.705151, -2.810553, -1.196685, 1.570796, 1.570748],accel_mss,speed_ms,0,blend_radius_m)
  movel([-0.010548, -0.706748, -2.810357, -1.195285, 1.570796, 1.560248],accel_mss,speed_ms,0,blend_radius_m)
  movel([-0.021606, -0.709535, -2.810011, -1.192843, 1.570796, 1.549190],accel_mss,speed_ms,0,blend_radius_m)
  movel([-0.033162, -0.713510, -2.809511, -1.189368, 1.570796, 1.537634],accel_mss,speed_ms,0,blend_radius_m)
  movel([-0.039102, -0.715945, -2.809202, -1.187242, 1.570796, 1.531694],accel_mss,speed_ms,0,blend_radius_m)
  movel([-0.051271, -0.721702, -2.808459, -1.182228, 1.570796, 1.519526],accel_mss,speed_ms,0,blend_radius_m)
  movel([-0.057482, -0.725024, -2.808024, -1.179341, 1.570796, 1.513315],accel_mss,speed_ms,0,blend_radius_m)
  movel([-0.070094, -0.732535, -2.807021, -1.172833, 1.570796, 1.500702],accel_mss,speed_ms,0,blend_radius_m)
  movel([-0.078788, -0.738403, -2.806220, -1.167766, 1.570796, 1.492008],accel_mss,speed_ms,0,blend_radius_m)
  movel([-0.087499, -0.744976, -2.805303, -1.162110, 1.570796, 1.483298],accel_mss,speed_ms,0,blend_radius_m)
  movel([-0.096132, -0.752178, -2.804274, -1.155937, 1.570796, 1.474664],accel_mss,speed_ms,0,blend_radius_m)
  movel([-0.104601, -0.759948, -2.803137, -1.149304, 1.570796, 1.466195],accel_mss,speed_ms,0,blend_radius_m)
  movel([-0.112827, -0.768224, -2.801894, -1.142272, 1.570796, 1.457969],accel_mss,speed_ms,0,blend_radius_m)
  movel([-0.120726, -0.776934, -2.800549, -1.134906, 1.570796, 1.450070],accel_mss,speed_ms,0,blend_radius_m)
  movel([-0.128222, -0.786018, -2.799106, -1.127265, 1.570796, 1.442574],accel_mss,speed_ms,0,blend_radius_m)
  movel([-0.135243, -0.795411, -2.797570, -1.119408, 1.570796, 1.435553],accel_mss,speed_ms,0,blend_radius_m)
